PROGRAM MAIN
// =============================================================
// TEST RUCHU TRANSPORTEROW
// =============================================================
//
// Proba na maszynie: jedna paleta idzie trasa, w kazdym kroku
// pracuje PARA transporterow - ten, z ktorego paleta zjezdza,
// i ten, na ktory wjezdza.
//
// -------------------------------------------------------------
// CZUJNIKI
// -------------------------------------------------------------
// Podpiete czujniki koncza przejazd zamiast czasowki.
//
//   xUseSensors   = FALSE  wracamy na same czasowki, jak dotad
//   xStepWatchdog = FALSE  krok czeka na czujnik BEZ KONCA
//
// Na czas recznego wyzwalania czujnikow watchdog jest WYLACZONY:
// zaden krok nie przeskoczy sam, dopoki nie podasz sygnalu.
// Po podpieciu prawdziwych czujnikow warto go wlaczyc - wtedy
// martwy czujnik nie zatrzyma proby, tylko zglosi sie sam przez
// xStepTimeout i licznik nTimeouts.
//
// Kroki konczone czujnikiem:
//   st.2 -> st.3    IN2      st.7 -> st.8    IN7
//   st.3 -> st.4    IN3/IN4  st.8 -> st.11   IN8
//   st.6 -> st.7    IN5      st.12-> st.13   IN6
//   st.15-> st.16   IN10
//
// STACJA 1 nie ma czujnika w tej probie. Zamiast niego dziala
// bit xSt01_StackReady: TRUE = stoi tam stos i mozna nim jechac,
// zbocze 0 -> 1 = przyjechal nowy stos (licznik nStacksSeen).
//
// STACJA 4 bada JADACA palete - patrz ACT_MoveSt04.
//
// Wyjatkiem jest przejazd poprzeczny 8 -> 10: tam paleta lezy
// na lancuchu, rolki stacji 8 i 10 sa opuszczone i MUSZA stac.
// Jedzie sam falownik 7, przez tChainTime.
//
// -------------------------------------------------------------
// CO NIE JEST URUCHAMIANE
// -------------------------------------------------------------
// Falowniki 1, 2 i 3 sa ZABLOKOWANE w axDriveEnabled:
//   1  krzywka desztaplarki   - mechanika niegotowa
//   2  krzywka na stacji 8    - mechanika niegotowa
//   3  rolki dociskowe st. 4  - to nie jest transporter
//
// Blokada dziala niezaleznie od tabeli krokow: nawet gdyby
// krok zazadal takiego napedu, nie ruszy. Zeby go dopuscic,
// trzeba swiadomie ustawic bit w axDriveEnabled.
//
// -------------------------------------------------------------
// STEROWANIE
// -------------------------------------------------------------
//   START_TEST = TRUE   symulacja ruchu jedzie
//   START_TEST = FALSE  wszystkie napedy staja
//
//   xCmdResetDrives     kasuje bledy wszystkich falownikow,
//                       dziala na zbocze i sam sie zdejmuje
//
// Po wcisnieciu START maszyna sama sprawdza, czy ktorys naped
// nie stoi w bledzie, i probuje go skasowac - zanim cokolwiek
// ruszy. Jesli sie nie uda, zapala sie xResetFailed.
//
// Pelna aplikacja siedzi w PRG_Machine i na razie nie jest
// wywolywana.
VAR

	// =========================================================
	// STEROWANIE
	// =========================================================

	// GLOWNY BIT TESTU TRASY. TRUE = jedziemy, FALSE = stop.
	START_TEST			: BOOL;


	// =========================================================
	// PROBA CALOSCIOWA: DOWOZ -> DESZTAPLOWANIE -> STACJA 4
	// =========================================================
	//
	// Niezalezna od START_TEST. Wozi palety ze stacji 1 do
	// desztaplarki, potem kazda zwolniona palete przez stacje 4
	// z testem dociskow i ZATRZYMUJE ja na koncu stacji 4.
	// Palete zabiera sie stamtad recznie.

	// Potwierdzenie operatora: palety leza na stacji 1.
	// Kod sam go zdejmuje po przyjeciu - kolejny stos wymaga
	// podania go od nowa.
	xSt01_StackReady	: BOOL;

	// Start dowozu i obslugi transportu w tej probie
	START_FEED			: BOOL;

	// Ile palet przeszlo przez stacje 4
	nFeedPallets		: UDINT;

	// Podglad
	nFeedStep			: INT;
	sFeedPhase			: STRING(79);

	// Wewnetrzne sekwencji dowozu
	nFeedStepOld		: INT;
	xFeedNewStep		: BOOL;
	xFeedArmed			: BOOL;
	xFeedAdvance		: BOOL;
	tFeedStep			: TIME;
	tonFeedStep			: TON;
	rtrgFeedStart		: R_TRIG;

	// =========================================================
	// TOR WYJSCIOWY - DRUGA PALETA W MASZYNIE
	// =========================================================
	//
	// Transport jest rozbity na DWA niezalezne tory:
	//
	//   nFeedStep  tor A: stacja 1 -> 3 -> 4 -> cykl stacji 5
	//   nOutStep   tor B: stacja 5 -> 6 -> ... -> 16
	//
	// Dzieki temu paleta po rozrywaniu jedzie w strone stacji 16
	// SAMA, a desztaplarka moze w tym czasie wydac nastepna.
	// W maszynie sa wtedy dwie palety naraz.
	//
	// Zasob wspolny to transporter stacji 5 (naped 5) i blokada.
	// Dlatego tor A nie wjedzie na stacje 5, dopoki tor B z niej
	// nie zjedzie - patrz krok 75.
	//
	// nOutStep = 0 znaczy TOR B WOLNY.

	nOutStep			: INT;
	sOutPhase			: STRING(79);

	nOutStepOld			: INT;
	xOutNewStep			: BOOL;
	xOutArmed			: BOOL;
	xOutAdvance			: BOOL;
	tOutStep			: TIME;
	tonOutStep			: TON;

	// Stacja 5 skonczyla cykl i oddala palete torowi B.
	// Na tym sygnale desztaplarka wypuszcza nastepna palete.
	xSt05_Done			: BOOL;

	// Zadania startu torow. Tor URUCHAMIA SIE SAM, w swoim kroku 0.
	// Powod jest w komentarzu przy silniku krokow nizej - w skrocie:
	// krok wpisany z ZEWNATRZ wykonalby sie jeszcze w tym samym
	// cyklu, ze stara flaga xOutAdvance, i przeskoczylby natychmiast.
	// -----------------------------------------------------
	// STACJA 8 - POSADZENIE PALETY NOK NA LANCUCHU
	// -----------------------------------------------------
	//
	// Na stacji 8 nie ma blokady, a transporter chodzi tak
	// gladko, ze paleta zatrzymuje sie raz dalej, raz blizej.
	// Dlatego po tSt08_DropDelay od IN7 OPUSZCZAMY rolki: paleta
	// siada na lancuchu i to on ja wyhamowuje - zawsze tak samo.
	//
	// DOTYCZY WYLACZNIE PALET NOK, bo tylko one jada lancuchem.
	// Paleta OK jedzie dalej rolkami i zatrzymuje sie jak dotad -
	// dla niej nic sie nie zmienia.
	//
	// Dwie NIEZALEZNE czasowki od tego samego IN7:
	//   tFeedSt08Stop   zdjecie zadania z falownika (dobieg)
	//   tSt08_DropDelay opuszczenie rolek pod paleta
	tSt08_DropDelay		: TIME := T#830MS;
	tonSt08Drop			: TON;

	// Zatrzask: rolki stacji 8 maja zostac w dole, dopoki lancuch
	// nie zabierze palety. Bez niego kroki, ktore ich nie pisza,
	// podnosilyby je z powrotem.
	xSt08_RollDown		: BOOL;

	// Paleta jest na stacji 8 - od potwierdzenia IN7 do zabrania
	// jej przez lancuch. Na tej fladze chodzi tonSt08Drop, dzieki
	// czemu odliczanie NIE ZALEZY od tego, w ktorym kroku toru B2
	// paleta akurat stoi.
	xSt08_AtStation		: BOOL;

	// Czy TA paleta jedzie trasa odrzutu (lancuchem).
	// W tej probie wszystkie palety jada na stacje 16, wiec bit
	// jest TRUE. Gdy dojdzie klasyfikacja OK/NOK, ma go ustawiac
	// wynik badania, a nie operator.
	xSt08_PalletNOK		: BOOL := TRUE;

	xOutStart			: BOOL;
	xOut2Start			: BOOL;
	xOut3Start			: BOOL;

	// Droga ze stacji 5 wolna: tor B1 pusty i stacja 7 pusta
	xSt05_CanPass		: BOOL;

	// -----------------------------------------------------
	// BUFOROWANIE - TOR B ROZBITY NA TRZY ODCINKI
	// -----------------------------------------------------
	//
	// Odcinki wyznaczaja CZUJNIKI, bo tylko one wiedza, gdzie
	// naprawde stoi paleta:
	//
	//   nOutStep   B1  st.5 -> 6 -> 7    konczy sie na IN5
	//   nOut2Step  B2  st.7 -> 8         konczy sie na IN7
	//   nOut3Step  B3  st.8 -> ... -> 16 konczy sie na IN10
	//
	// Kazdy odcinek zwalnia sie DOPIERO wtedy, gdy nastepny
	// przejmie palete. Dzieki temu w obiegu moga byc naraz:
	// paleta na stacji 5, paleta na 7, paleta na 8 i paleta
	// w drodze na 16 - zamiast jednej na cala maszyne.
	//
	// Transporter stacji 7 (naped 11) obsluguje B1 i B2, a rolki
	// stacji 8 (naped 12) B2. Dlatego paleta czeka w krokach
	// 205 i 218 z ZATRZYMANYMI napedami, zamiast dojezdzac
	// wprost na zajety odcinek.

	nOut2Step			: INT;
	sOut2Phase			: STRING(79);
	nOut2StepOld		: INT;
	xOut2NewStep		: BOOL;
	xOut2Armed			: BOOL;
	xOut2Advance		: BOOL;
	tOut2Step			: TIME;
	tonOut2Step			: TON;

	nOut3Step			: INT;
	sOut3Phase			: STRING(79);
	nOut3StepOld		: INT;
	xOut3NewStep		: BOOL;
	xOut3Armed			: BOOL;
	xOut3Advance		: BOOL;
	tOut3Step			: TIME;
	tonOut3Step			: TON;

	// -----------------------------------------------------
	// STACJA 5 - CZAS PCHANIA PALETY DO BLOKADY
	// -----------------------------------------------------
	//
	// Paleta opiera sie o blokade duzo wczesniej, niz konczy sie
	// krok 80. Kazda sekunda ponad to jest transporterem
	// mielacym pod stojaca paleta - tak przeciazamy naped 5.
	// Po tym czasie napedy 4 i 5 STAJA, a krok trwa dalej.
	//
	// DOMYSLNIE ROWNE tFeedToSt05 - czyli tak, jak bylo przed
	// wprowadzeniem tej nastawy. Moje 4 s bylo za krotkie
	// i paleta nie dojezdzala do blokady.
	//
	// Skracaj DOPIERO po obejrzeniu, gdzie paleta sie zatrzymuje:
	// ma byc na tyle dlugie, zeby doszla do blokady, i na tyle
	// krotkie, zeby transporter nie mielil pod nia bez potrzeby.
	tSt05_Push			: TIME := T#9S;
	tonSt05Push			: TON;

	// -----------------------------------------------------
	// STACJA 4 - ROLKI DOCISKOWE (NAPED 3)
	// -----------------------------------------------------
	//
	// Kreca sie razem z transporterem stacji 4 (naped 4).
	// Bit ponizej wybiera kierunek obrotu - do ustawienia
	// online, bez pobierania projektu.
	xSt04_RollRev		: BOOL := TRUE;

	// Stan dociskow stacji 4 w tej probie - przepisywany co cykl
	xFeedPressOn		: BOOL;
	xFeedPressLoOn		: BOOL;

	// Czas przejazdu st.4 -> st.5. Stacja 5 nie ma czujnika,
	// wiec dojazd konczy sie czasowka. Dobrane na maszynie.
	tFeedToSt05			: TIME := T#9S;

	// DOBIEG NA STACJI 3. Czujnik IN2 widzi krawedz natarcia
	// stosu, a szczeki maja trafic pod DRUGA palete od dolu -
	// stos musi wiec dojechac jeszcze kawalek po wykryciu.
	//
	// ZERO = stop natychmiast po czujniku, czyli tak, jak bylo.
	// Odpowiednik tSt04_StopDelay dla stacji 4.
	tFeedSt03Stop		: TIME := T#0S;

	// Odstep od zatrzymania palety na stacji 5 do ruszenia
	// mechaniki. Stacja 5 nie ma czujnika, wiec nie wiemy, kiedy
	// paleta oprze sie o blokade - dajemy jej na to czas.
	tSt05_Settle		: TIME := T#8S;

	// Stan mechaniki stacji 5 w tej probie - kazdy krok podaje
	// swoj pelny stan, cewki przepisujemy co cykl.
	xFeed05_Block		: BOOL;		// blokada wysunieta
	xFeed05_Lift		: BOOL;		// szczeki podniesione
	xFeed05_Jaws		: BOOL;		// szczeki zamkniete
	xFeed05_Pull		: BOOL;		// silowniki rozrywajace w gorze

	// Diagnostyka napedow zadanych przez biezacy krok
	nFeedBadDrv			: INT;
	sFeedDrvWhy			: STRING(31);
	tonFeedDrv			: TON;

	// -----------------------------------------------------
	// CZASOWKI PRZEJAZDOW BEZ CZUJNIKA
	// -----------------------------------------------------
	//
	// Odcinki, na ktorych nie ma czym potwierdzic dojazdu.
	// Tam, gdzie czujnik jest, czasowka nie jest uzywana wcale.

	tFeed5to6			: TIME := T#12S;		// st.5 -> st.6
	tFeed9Chain			: TIME := T#19S;		// lancuch st.8 -> st.10
	tFeed10to14			: TIME := T#8S;		// st.10 -> st.14
	tFeed14to15			: TIME := T#8S;		// st.14 -> st.15

	// Paleta zniknela z czujnika stacji 16. Po tym czasie
	// uznajemy stacje za pusta - odbiera ja operator.
	tSt16_Clear			: TIME := T#4S;

	// -----------------------------------------------------
	// DOBIEGI PO CZUJNIKACH
	// -----------------------------------------------------
	//
	// Czujnik widzi krawedz natarcia palety, a ona ma stanac
	// na srodku stacji. ZERO = stop natychmiast po czujniku.
	// Odpowiedniki tFeedSt03Stop i tSt04_StopDelay.

	tFeedSt08Stop		: TIME := T#740MS;		// IN7  stacja 8
	tFeedSt16Stop		: TIME := T#0S;		// IN10 stacja 16

	// Rolki podnoszone stacji 8 i 10. TRUE = w gorze, czyli
	// transport wzdluz. Na czas przejazdu lancuchem OBIE musza
	// zejsc, inaczej szarpalyby palete z dwoch stron.
	xFeedRoll08Up		: BOOL := TRUE;
	xFeedRoll10Up		: BOOL := TRUE;

	// Zezwolenie z lancucha bezpieczenstwa
	xSafetyOK			: BOOL := TRUE;

	// KASOWANIE BLEDOW WSZYSTKICH FALOWNIKOW - dziala na zbocze.
	// Bit sam sie zdejmuje po wystawieniu impulsu.
	xCmdResetDrives		: BOOL;

	// Automatyczne kasowanie bledow po wcisnieciu START.
	// FALSE = start nie probuje niczego kasowac.
	xAutoResetOnStart	: BOOL := TRUE;

	// Odstep miedzy kolejnymi probami kasowania
	tResetGap			: TIME := T#1S;

	// Czestotliwosc BAZOWA transporterow [Hz]. Uzywana wszedzie,
	// gdzie alrDriveFreq nie ma wpisanej wlasnej wartosci.
	lrTestFreq			: LREAL := 20.0;

	// =========================================================
	// CZESTOTLIWOSC OSOBNO DLA KAZDEGO NAPEDU [Hz]
	// =========================================================
	//
	// Zero znaczy "uzyj lrTestFreq". Wpisanie liczby dotyczy
	// tylko tego jednego falownika.
	//
	// Przydzial stacja -> falownik:
	//   st.1  -> 8     st.5  -> 5     st.9  -> 7      st.13 -> 15
	//   st.2  -> 9     st.6  -> 6     st.10 -> 16     st.14 -> 17
	//   st.3  -> 10    st.7  -> 11    st.11 -> 13     st.15 -> 18
	//   st.4  -> 4     st.8  -> 12    st.12 -> 14     st.16 -> 19
	//
	// Krzywki 1 i 2 maja wlasna lrCamFreq i ta tablica ich nie
	// dotyczy.
	//
	// UWAGA: naped czyta czestotliwosc przy STARCIE (M_Start jest
	// wolane na zboczu). Zmiana w trakcie jazdy zadziala dopiero
	// przy nastepnym ruszeniu.

	alrDriveFreq		: ARRAY[1..20] OF LREAL;

	// Czas jednego kroku - przejazd palety miedzy stacjami
	tStepTime			: TIME := T#5S;

	// Przejazd poprzeczny transporterem lancuchowym jest dluzszy
	tChainTime			: TIME := T#6S;

	// Czas jednego ruchu silownika. Czujnikow polozenia jeszcze
	// nie ma, wiec po tym czasie uznajemy ruch za wykonany.
	tCylTime			: TIME := T#2S;

	// Stacja 4 - dociski gorne i dolne maja isc praktycznie razem.
	// Gorne schodza pierwsze, dolne po tym krotkim odstepie,
	// zeby dolne nie uniosly palety. Cofanie jest jednoczesne.
	tSt04_UpToLo		: TIME := T#2200MS;

	// FALSE = same transportery, silowniki stoja
	xCylEnable			: BOOL := TRUE;


	// =========================================================
	// CZUJNIKI
	// =========================================================
	//
	// FALSE = jedziemy na samych czasowkach, tak jak dotad.
	// TRUE  = kroki wypisane w ACT_Move koncza sie czujnikiem,
	//         a czasowka pracuje juz tylko jako watchdog.

	xUseSensors			: BOOL := TRUE;

	// STACJA 1 - czujnika IN1 NIE uzywamy. Zastepuje go bit
	// xSt01_StackReady zadeklarowany na gorze.
	nStacksSeen			: UDINT;

	// Obraz czujnikow sprowadzony do JEDNEGO znaczenia:
	// TRUE = PALETA JEST. Polaryzacje ustawia ACT_Inputs i tylko on.
	xPal_St03			: BOOL;		// IN2   stacja 3
	xPal_St04In			: BOOL;		// IN3   wjazd na stacje 4
	xPal_St04End		: BOOL;		// IN4   koniec testu desek
	xPal_St07			: BOOL;		// IN5   stacja 7
	xPal_St13			: BOOL;		// IN6   koniec stacji 13
	xPal_St08			: BOOL;		// IN7   stacja 8
	xPal_St11			: BOOL;		// IN8   stacja 11
	xPal_St16			: BOOL;		// IN10  stacja 16

	// Surowe wejscia - do podgladu bez otwierania GVL
	axInRaw				: ARRAY[1..10] OF BOOL;

	// -----------------------------------------------------
	// POLARYZACJA CZUJNIKOW - JEDYNE MIEJSCE
	// -----------------------------------------------------
	//
	// TRUE  = czujnik ROZWIERA przy palecie (0 = paleta)
	// FALSE = czujnik ZWIERA przy palecie   (1 = paleta)
	//
	// Wartosci ponizej sa wg opisu z maszyny. Jesli ktorys
	// czujnik zachowa sie odwrotnie, przestawia sie JEDEN bit
	// online - bez zmiany kodu i bez pobierania projektu.
	//
	//   1  st.1              nieuzywany
	//   2  st.3              ROZWIERA - stwierdzone na maszynie,
	//                        wbrew pierwotnemu opisu
	//   3  wjazd st.4        rozwiera
	//   4  koniec testu st.4 rozwiera
	//   5  st.7              zwiera
	//   6  koniec st.13      rozwiera
	//   7  st.8              zwiera
	//   8  st.11             zwiera
	//   9  niepodlaczony
	//  10  st.16             zwiera

	axInInverted		: ARRAY[1..10] OF BOOL :=
	                      [FALSE, TRUE, TRUE, TRUE, FALSE,
	                       TRUE, FALSE, FALSE, FALSE, FALSE];

	// WATCHDOG KROKU CZUJNIKOWEGO.
	//
	// FALSE = krok czeka na czujnik BEZ KONCA. Tak jedziemy przy
	//         recznym wyzwalaniu czujnikow - nic nie przeskoczy
	//         kroku, dopoki sam nie podasz sygnalu.
	// TRUE  = po tMoveTimeout krok konczy sie mimo wszystko,
	//         zapala sie xStepTimeout i rosnie nTimeouts.
	xStepWatchdog		: BOOL := FALSE;

	tMoveTimeout		: TIME := T#20S;
	xStepTimeout		: BOOL;
	nTimeouts			: UDINT;


	// =========================================================
	// STACJA 4 - TEST NA JADACEJ PALECIE
	// =========================================================
	//
	// Paleta nie zatrzymuje sie pod rolkami. Czujnik wjazdu (IN3)
	// odlicza tSt04_EntryToPress i wtedy rolki schodza na deski.
	// Czujnik konca testu (IN4) NATYCHMIAST je cofa, a transporter
	// stoi tSt04_StopDelay pozniej - paleta dojezdza do konca stacji.

	tSt04_EntryToPress	: TIME := T#2600MS;
	tSt04_StopDelay		: TIME := T#300MS;


	// =========================================================
	// SZTAPLARKA I DESZTAPLARKA
	// =========================================================
	//
	// Dwa NIEZALEZNE cykle, kazdy z wlasnym bitem startu. Nie
	// maja nic wspolnego z START_TEST.
	//
	// Poziom TRUE = cykl pracuje.
	// Poziom FALSE = natychmiastowy stop, hamulec zaklada sie
	//                tCamBrakeHold pozniej.
	//
	// REGULA NADRZEDNA obu maszyn: nic w szczekach = szczeki
	// OTWARTE i jazda na pozycje DOLNA, niezaleznie od tego,
	// gdzie wozek stoi. Cykl zaczyna sie i konczy na dole
	// z otwartymi szczekami.

	START_DESTACK		: BOOL;		// desztaplarka, stacja 3
	START_STACK			: BOOL;		// sztaplarka, stacja 11

	// -----------------------------------------------------
	// JAZDA RECZNA KRZYWKA
	// -----------------------------------------------------
	//
	// Trzymasz bit - wozek jedzie. Puszczasz - staje, hamulec
	// zaklada sie tCamBrakeHold pozniej, tak samo jak w cyklu.
	//
	// Dziala TYLKO przy zdjetym starcie danej maszyny, zeby
	// nigdy nie walczyc z sekwencja. Sluzy do sprawdzenia,
	// czy enkoder liczy i w ktora strone.

	JOG_DESTACK_FWD		: BOOL;
	JOG_DESTACK_REV		: BOOL;
	JOG_STACK_FWD		: BOOL;
	JOG_STACK_REV		: BOOL;

	xDeJog				: BOOL;
	xStJog				: BOOL;

	// -----------------------------------------------------
	// UCZENIE POZYCJI
	// -----------------------------------------------------
	//
	// Dojedz jogiem tam, gdzie wozek ma stawac, i podaj bit.
	// Zbocze 0 -> 1 przepisuje BIEZACA pozycje enkodera do
	// odpowiedniej nastawy. Koniec z wpisywaniem liczb z palca.
	//
	// UWAGA: nastawy siedza na razie w MAIN, wiec pobranie
	// projektu je kasuje. Po ustaleniu przenosimy do GVL_PERSIST.

	TEACH_DE_BOTTOM		: BOOL;
	TEACH_DE_MIDDLE		: BOOL;
	TEACH_DE_TOP		: BOOL;
	TEACH_ST_BOTTOM		: BOOL;
	TEACH_ST_MIDDLE		: BOOL;
	TEACH_ST_TOP		: BOOL;

	rtrgTeach			: ARRAY[1..6] OF R_TRIG;

	// Ostatnio nauczona pozycja - potwierdzenie na podgladzie
	sTeachLast			: STRING(79);

	// Czestotliwosc krzywek. Osobno od transporterow.
	// Nizej niz transportery - wolniej znaczy krotszy dojazd
	// po zdjeciu zadania, a wiec mniejszy blad pozycji.
	lrCamFreq			: LREAL := 15.0;

	// Ruch szczek - czujnikow polozenia nie ma
	tJawTime			: TIME := T#2S;


	// Odstep od ZALOZENIA hamulca do chwytu szczekami.
	// Wozek musi sie uspokoic, zanim szczeki wejda pod palete.
	tDeGripDelay		: TIME := T#1S;

	// -----------------------------------------------------
	// POZYCJE I LICZNIKI SIEDZA W GVL_PERSIST
	// -----------------------------------------------------
	//
	// Nastawy:  GVL_PERSIST.St03.Cfg.diPosBottom / Middle / Top
	//           GVL_PERSIST.St11.Cfg.diPosBottom / Middle / Top
	//           GVL_PERSIST.St03.Cfg.nStackSize
	// Liczniki: GVL_PERSIST.St03.Mem.nRemaining / nHeld
	//           GVL_PERSIST.St11.Mem.nHeld
	//
	// Sa NIEULOTNE, wiec przezywaja zanik zasilania, aktywacje
	// konfiguracji i reset cold. Uczenie pozycji zapisuje wprost
	// tam - nie ma drugiej kopii, ktora moglaby sie rozjechac.



	// Wyprzedzenie hamowania - zadanie znika tyle przed celem.
	// Zaczynamy od zera i ustawiamy z odczytu diCoast.
	diCamStopLead		: DINT := 0;

	// Okno "jestem na miejscu" przy bazowaniu. Bez niego wozek
	// stojacy tuz przy dolnej pozycji robilby caly obrot, zeby
	// do niej "dojechac".
	diCamTol			: DINT := 300;

	// Ile impulsow za celem uznajemy jeszcze za "jestem".
	// Musi byc WIEKSZE niz dojazd po zdjeciu zadania, inaczej
	// wozek stojacy tuz ZA punktem objechalby caly obrot,
	// zeby do niego wrocic.
	diCamOvershoot		: DINT := 5000;

	// -----------------------------------------------------
	// DOKAD JEDZIE BIEZACY KROK
	// -----------------------------------------------------
	//
	// Krok podaje WARTOSC ENKODERA, do ktorej ma dojechac,
	// a droge liczymy raz, przy wejsciu w krok, z zywej
	// pozycji. Nigdzie nie zakladamy, ile impulsow ma cykl
	// maszyny - to bylo zrodlo kumulujacego sie bledu.

	diDeGoToEnc			: DINT;
	diStGoToEnc			: DINT;

	// -----------------------------------------------------
	// POMIAR - ILE IMPULSOW MA NAPRAWDE CYKL MASZYNY
	// -----------------------------------------------------
	//
	// diDeCycleCounts   droga przejechana miedzy kolejnymi
	//                   dolnymi pozycjami. Jesli enkoder jest
	//                   1:1 z korba, ma byc okolo 65536.
	//                   Kazda inna liczba znaczy, ze cykl
	//                   maszyny to nie jest jeden obrot enkodera.
	// diDeBottomErr     o ile minelismy nauczony dol, ze znakiem
	// diDeCoastMax      najwiekszy zaobserwowany dojazd. Musi
	//                   byc MNIEJSZY niz diCamOvershoot, inaczej
	//                   ruch do punktu tuz za nami pojedzie
	//                   dookola.

	diDeCycleCounts		: DINT;
	diDeBottomErr		: DINT;
	diDeCoastMax		: DINT;

	diStCycleCounts		: DINT;
	diStBottomErr		: DINT;
	diStCoastMax		: DINT;

	// Ustawienie punktu odniesienia osi, impuls jednocyklowy
	xDeSetAccum			: BOOL;
	xStSetAccum			: BOOL;
	diDeAccumSet		: DINT;
	diStAccumSet		: DINT;

	// Roboczy
	diTmp				: DINT;

	// -----------------------------------------------------
	// KONTROLA POPRAWNOSCI NASTAW POZYCJI
	// -----------------------------------------------------
	//
	// Trzy pozycje musza byc od siebie ODDALONE. Zerowe albo
	// pomylone nastawy oznaczaja, ze wozek "juz jest na miejscu"
	// w kazdym kroku - a wtedy szczeki zamykaja sie na dole,
	// na stosie. Cykl nie ma prawa ruszyc na takich nastawach.

	xDeCfgOK			: BOOL;
	xStCfgOK			: BOOL;
	diCamMinSpan		: DINT := 1000;

	// -----------------------------------------------------
	// KONTROLA ENKODERA PO STARCIE
	// -----------------------------------------------------
	//
	// Enkoder absolutny powinien utrzymac wartosc przez zanik
	// zasilania. Zapamietujemy ja na biezaco w GVL_PERSIST
	// i po starcie porownujemy z odczytem. Zgadza sie -
	// bazowanie jest zbedne. Nie zgadza sie - kod to zglasza,
	// zamiast po cichu jechac wedlug zlych pozycji.

	xEncCheckDone		: BOOL;
	diDeEncJump			: DINT;
	diStEncJump			: DINT;
	sEncCheck			: STRING(79);

	// Ile impulsow roznicy jeszcze wybaczamy po starcie
	diEncCheckTol		: DINT := 500;

	// START: wyprzedzenie zdjecia hamulca przed komenda dla
	// falownika. ZERO = jednoczesnie, i tak ma byc.
	tCamBrakeRelease	: TIME := T#0S;

	// STOP: ile hamulec czeka po zdjeciu komendy z falownika.
	// Rampa hamowania falownika to 1 s, wiec hamulec zaciska sie
	// na wolno obracajacym sie jeszcze wale - SWIADOMIE, zeby
	// nie puszczac wozka wolno.
	tCamBrakeHold		: TIME := T#700MS;

	// Kasowanie czuwaka obu osi, dziala na zbocze
	RESET_CAM			: BOOL;

	// =========================================================
	// RESET CYKLU DO ZERA
	// =========================================================
	//
	// Po recznym oproznieniu maszyny z palet. Sprowadza obie
	// maszyny i transport do kroku 0, zeruje liczniki palet
	// i uzgodnienia, kasuje czuwaki osi.
	//
	// NICZYM NIE RUSZA. Wozki wroca na dol dopiero przy starcie,
	// bo krok 0 obu maszyn to "szczeki otwarte, jazda na dol".
	//
	// Bit sam sie zdejmuje.

	RESET_CYCLE			: BOOL;
	rtrgResetCycle		: R_TRIG;

	// -----------------------------------------------------
	// PODGLAD OSI
	// -----------------------------------------------------

	fbCamDestack		: FB_CamAxis;
	fbCamStack			: FB_CamAxis;

	nDeStep				: INT;
	nStStep				: INT;
	sDePhase			: STRING(79);
	sStPhase			: STRING(79);
	nDeCycles			: UDINT;
	nStCycles			: UDINT;

	// -----------------------------------------------------
	// LICZNIKI PALET
	// -----------------------------------------------------
	//
	// GVL_PERSIST.St03.Mem.nRemaining  ile palet zostalo w desztaplarce razem:
	//               na transporterze plus wiszace na szczekach
	// GVL_PERSIST.St03.Mem.nHeld       ile wisi na szczekach desztaplarki
	// GVL_PERSIST.St11.Mem.nHeld       ile palet liczy stos w sztaplarce


	// -----------------------------------------------------
	// UZGODNIENIA Z TRANSPORTEM
	// -----------------------------------------------------

	// Desztaplarka zwolnila palete - transport moze ja zabrac
	xDe_PalletReleased	: BOOL;

	// Desztaplarka pusta, cykl zamkniety na pozycji dolnej
	xDe_Empty			: BOOL;

	// Sztaplarka ma pelny stos na transporterze
	xSt_StackReady		: BOOL;

	// -----------------------------------------------------
	// CZASOWKI OD ZALOZENIA HAMULCA
	// -----------------------------------------------------
	//
	// Licza dopiero od chwili, w ktorej hamulec sie ZACISNIE -
	// nie od wejscia w krok.

	tonDeBrake			: TON;
	tonStBrake			: TON;
	tDeBrakeWait		: TIME;
	tStBrakeWait		: TIME;

	// Czujnik musi byc najpierw WOLNY, zeby sie zaliczyl
	xDeArmed			: BOOL;
	xStArmed			: BOOL;

	// Stan szczek deklarowany przez KAZDY krok i przepisywany
	// na cewki co cykl. Poleganie na tym, ze cewka zachowa
	// wartosc miedzy krokami, juz raz nas kosztowalo prawdziwy
	// blad - ACT_ClearCoils zeruje je w kazdym cyklu.
	xDeJawsClosed		: BOOL;
	xStJawsClosed		: BOOL;

	// -----------------------------------------------------
	// ZYCIE ENKODEROW
	// -----------------------------------------------------
	//
	// Rosna przy KAZDEJ zmianie pozycji. Jesli silnik chodzi,
	// a licznik stoi - enkoder nie jest podlinkowany albo nie
	// liczy. To rozstrzyga sprawe w jednej liczbie.

	nDeEncMoves			: UDINT;
	nStEncMoves			: UDINT;
	diDePosOld			: DINT;
	diStPosOld			: DINT;

	tonDeStep			: TON;
	tonStStep			: TON;
	xDeAdvance			: BOOL;
	xStAdvance			: BOOL;
	tDeStep				: TIME;
	tStStep				: TIME;

	// Zadanie dla osi - liczone przez maszyne stanow,
	// podawane do bloku JEDNYM wywolaniem na cykl
	xDeGo				: BOOL;
	xStGo				: BOOL;
	diDeTarget			: DINT;
	diStTarget			: DINT;

	// Wykrycie zmiany kroku. Bez tego krok zaliczylby xInPos
	// z POPRZEDNIEJ pozycji i przeskoczyl dwa kroki naraz.
	nDeStepOld			: INT;
	nStStepOld			: INT;
	xDeNewStep			: BOOL;
	xStNewStep			: BOOL;
	xDeAtPos			: BOOL;
	xStAtPos			: BOOL;

	rtrgDeStart			: R_TRIG;
	rtrgStStart			: R_TRIG;

	// Cewki hamulcow. TRUE = hamulec ROZLACZONY.
	xBrakeDestack		: BOOL;
	xBrakeStack			: BOOL;


	// =========================================================
	// RECZNE STEROWANIE POJEDYNCZYM SILOWNIKIEM
	// =========================================================
	//
	// Do sprawdzenia okablowania bez sekwencji. Gdy nManCyl <> 0,
	// sekwencja stoi, transportery stoja, a wybrany silownik
	// slucha bitow ponizej.
	//
	//    1  st.3  szczeki desztaplarki
	//    2  st.4  dociski gorne
	//    3  st.4  dociski dolne
	//    4  st.5  blokada
	//    5  st.5  podnoszenie szczek
	//    6  st.5  szczeki (zamkniecie / otwarcie)
	//    7..12 st.5 silowniki rozrywajace 1..6
	//   13  st.8  rolki podnoszone
	//   14  st.10 rolki podnoszone
	//   15  st.11 szczeki sztaplarki

	nManCyl				: INT;
	xManExtend			: BOOL;
	xManRetract			: BOOL;


	// =========================================================
	// DOPUSZCZENIE NAPEDOW
	// =========================================================
	//
	// FALSE = naped nie ruszy, chocby krok tego zadal.
	// Ustawiane w ACT_Config, mozna zmieniac online.

	axDriveEnabled		: ARRAY[1..20] OF BOOL;


	// =========================================================
	// KIERUNEK OBROTOW
	// =========================================================
	//
	// TRUE = jazda w druga strone. Silniki stacji 1, 5, 6, 7,
	// 8, 9, 14, 15, 16 sa podlaczone odwrotnie - do poprawy
	// w szafie, na razie odwracamy bit.

	axReverse			: ARRAY[1..20] OF BOOL;


	// =========================================================
	// PODGLAD
	// =========================================================

	// Gdzie jest wirtualna paleta i co sie z nia dzieje
	nIdx				: INT;		// pozycja na trasie
	nSub				: INT;		// krok sekwencji stacji
	xMoving				: BOOL;		// TRUE = przejazd, FALSE = praca stacji
	sPhase				: STRING(79);

	// Ktore napedy maja teraz pracowac
	axRunReq			: ARRAY[1..20] OF BOOL;

	// Stan napedow
	aeDrvState			: ARRAY[1..20] OF E_NordSK550P_State;
	axDrvRunning		: ARRAY[1..20] OF BOOL;
	alrDrvFreqAct		: ARRAY[1..20] OF LREAL;

	// UWAGA - to sa DWIE ROZNE rzeczy:
	//   axDrvFault  blad zglaszany przez falownik (bit 3 StatusWord)
	//   axDrvError  jakakolwiek blokada: blad, brak zezwolenia
	//               albo zerwana komunikacja
	axDrvFault			: ARRAY[1..20] OF BOOL;
	axDrvError			: ARRAY[1..20] OF BOOL;

	// Slowa sterujace i statusowe - do czytania, co naped
	// naprawde zglasza
	awDrvStatus			: ARRAY[1..20] OF UINT;
	awDrvControl		: ARRAY[1..20] OF UINT;

	// Ktorykolwiek naped zglasza blad
	xAnyDriveError		: BOOL;
	xAnyDriveFault		: BOOL;

	// Kasowanie nie poskutkowalo - blad wraca albo trzyma
	xResetFailed		: BOOL;

	// Trwa kasowanie bledow przed startem
	xResetInProgress	: BOOL;
	nResetTries			: INT;

	// Blokada zadzialala - lancuch wymusil postoj rolek 8 i 10
	xChainInterlock		: BOOL;

	// Blokada stacji 5 kontra transporter - patrz ACT_ApplyDrives
	xSt05_BlockLock		: BOOL;
	tonSt05BlockDown	: TON;

	// Czas biezacego kroku
	tThisStep			: TIME;

	// Licznik pelnych przebiegow trasy
	nLoops				: UDINT;

	// =========================================================
	// LICZNIKI ZYCIA - do sprawdzenia, co sie naprawde wykonuje
	// =========================================================
	//
	// nCycles     rosnie w kazdym cyklu zadania. Jesli stoi,
	//             MAIN sie nie wykonuje albo wysypal sie wczesniej.
	// nOutWrites  rosnie za kazdym przepisaniem cewek na wyjscia.
	//             Jesli nCycles rosnie, a nOutWrites stoi -
	//             program nie dochodzi do ACT_Outputs.
	// nCoilsOn    ile cewek jest w tej chwili podanych. Jesli
	//             rosnie i spada, a nic sie nie rusza - sygnal
	//             nie dochodzi do zaworu.

	nCycles				: UDINT;
	nOutWrites			: UDINT;
	nCoilsOn			: INT;


	// =========================================================
	// CEWKI ZAWOROW
	// =========================================================
	//
	// Stan trzymany miedzy cyklami. ACT_Outputs przepisuje go
	// na wyjscia - mapowanie jest TAM i tylko tam.

	// Stacja 3 - szczeki desztaplarki
	xSt03_JawClose		: BOOL;
	xSt03_JawOpen		: BOOL;

	// Stacja 4 - dociski. Obie grupy gornych chodza razem.
	xSt04_UpExt			: BOOL;
	xSt04_UpRet			: BOOL;
	xSt04_LoExt			: BOOL;
	xSt04_LoRet			: BOOL;

	// Stacja 5
	xSt05_BlockExt		: BOOL;		// blokada wysuw
	xSt05_BlockRet		: BOOL;		// blokada opuszczenie
	xSt05_LiftUp		: BOOL;		// szczeki w gore
	xSt05_LiftDown		: BOOL;		// szczeki w dol
	xSt05_JawClose		: BOOL;		// trzy pary szczek razem
	axSt05_PullUp		: ARRAY[1..6] OF BOOL;
	axSt05_PullDown		: ARRAY[1..6] OF BOOL;

	// Rolki podnoszone
	xSt08_Up			: BOOL;
	xSt08_Down			: BOOL;
	xSt10_Up			: BOOL;
	xSt10_Down			: BOOL;

	// Stacja 11 - szczeki sztaplarki
	xSt11_JawClose		: BOOL;
	xSt11_JawOpen		: BOOL;


	// =========================================================
	// NAPEDY
	// =========================================================

	fbNord				: ARRAY[1..20] OF FB_NordSK550PP;


	// =========================================================
	// OBSERWATOR STANU - LOG CSV NA DYSKU STEROWNIKA
	// =========================================================
	//
	// Co tLogPeriod jeden wiersz z kluczowymi zmiennymi, a do
	// tego wiersz na kazde ZDARZENIE: zmiana numeru kroku,
	// czujnika, zadania napedu, bledu falownika, bitu operatora,
	// szczek, skok enkodera. Najwyzej jeden wiersz na cykl.
	//
	// Nowy plik: start PLC, RESET_CYCLE, zbocze xLogNewFile.
	// Katalog MUSI istniec na sterowniku: fbLog.sDir
	// (domyslnie C:\TesterPalet\log\). Nazwa pliku w fbLog.sFileName.
	//
	// Logger tylko CZYTA zmienne procesu - ACT_Logger idzie jako
	// ostatnia akcja cyklu, po ACT_Outputs, zeby w pliku bylo to,
	// co naprawde poszlo na wyjscia.

	fbLog				: FB_CsvLogger;

	// FALSE = nie zbieramy wierszy (plik zostaje, nic sie nie psuje)
	xLogEnable			: BOOL := TRUE;

	// Zbocze = nowy plik bez resetu cyklu. Sam sie zdejmuje.
	xLogNewFile			: BOOL;

	// Takt wiersza okresowego
	tLogPeriod			: TIME := T#1S;
	tonLog				: TON;

	// Skok enkodera w jednym cyklu, od ktorego piszemy zdarzenie
	diLogEncJump		: DINT := 2000;

	// Powod biezacego wiersza - do kolumny "why"
	sLogWhy				: STRING(79);
	xLogEvent			: BOOL;
	nLogRows			: UDINT;

	// Pamiec do wykrywania zdarzen
	xLogInit			: BOOL;
	anLogStepOld		: ARRAY[1..6] OF INT;
	axLogInOld			: ARRAY[1..10] OF BOOL;
	axLogReqOld			: ARRAY[1..20] OF BOOL;
	axLogFaultOld		: ARRAY[1..20] OF BOOL;
	axLogBitOld			: ARRAY[1..24] OF BOOL;
	axLogBit			: ARRAY[1..24] OF BOOL;

	// Robocze do skladania nazw kolumn napedow
	sLogPfx				: STRING(15);
	wLogFesto1			: WORD;
	wLogFesto2			: WORD;
	nLogI				: INT;
	nLogJ				: INT;


	// =========================================================
	// WEWNETRZNE
	// =========================================================

	xInit				: BOOL;
	i					: INT;
	lrThisFreq			: LREAL;
	tonStep				: TON;
	tonResetGap			: TON;
	xAdvance			: BOOL;
	rtrgStart			: R_TRIG;
	rtrgResetDrv		: R_TRIG;
	rtrgStack			: R_TRIG;
	xDoResetPulse		: BOOL;
	axRunOld			: ARRAY[1..20] OF BOOL;

	// Krok zglasza tu, ze czeka na czujnik i ktory to czujnik.
	// Kasowane co cykl, ustawiane przez sam krok.
	xWaitSensor			: BOOL;
	xSensorOK			: BOOL;

	// Czujnik musi najpierw byc WOLNY. Bez tego zaliczylby sie
	// stan sprzed kroku albo czujnik zawieszony na stale.
	xStepArmed			: BOOL;

	// Wykrycie zmiany kroku - czasowka i uzbrojenie od zera
	xNewStep			: BOOL;
	nIdxOld				: INT;
	nSubOld				: INT;
	xMovingOld			: BOOL;

	// TRUE = przejazd ma jeszcze kroki wewnetrzne, nIdx zostaje
	xHoldIdx			: BOOL;

END_VAR
VAR CONSTANT

	// P105 falownikow
	cFmax				: LREAL := 50.0;

	// Liczba falownikow zmapowanych w .tsproj
	cNumDrives			: INT := 19;

	// Liczba pozycji na trasie
	cLastIdx			: INT := 16;

	// Ile razy probujemy skasowac blad przed startem
	cResetTries			: INT := 3;

END_VAR

// =============================================================
// MAIN - TEST RUCHU TRANSPORTEROW
// =============================================================

// Puls zycia - jesli ten licznik stoi, MAIN sie nie wykonuje
nCycles := nCycles + 1;

ACT_Config();

ACT_Inputs();

ACT_Sequence();

// Krzywki chodza NIEZALEZNIE od START_TEST i po ACT_Sequence,
// zeby ich szczeki mialy pierwszenstwo przed sekwencja linii.
ACT_CamCycles();

// Transport proby calosciowej - po krzywkach, zeby jego
// cewki i zadania napedow mialy pierwszenstwo.
ACT_TestFeed();

ACT_ResetDrives();

ACT_ApplyDrives();

ACT_Drives();

ACT_Outputs();

// Obserwator stanu - OSTATNI, zeby logowal to, co poszlo na wyjscia
ACT_Logger();

ACTION ACT_ApplyDrives:
// =============================================================
// ACT_ApplyDrives
// Zadanie ruchu -> metody falownikow
// =============================================================
//
// Metody wolamy NA ZBOCZU. Blok napedu przy blokadzie sam kasuje
// zadanie ruchu i naped nie moze ruszyc sam po ustapieniu
// przyczyny - wolanie M_Start co cykl zepsuloby to zabezpieczenie.

xAnyDriveError := FALSE;


// -------------------------------------------------------------
// BLOKADA: LANCUCH KONTRA ROLKI STACJI 8 I 10
// -------------------------------------------------------------
//
// Gdy jedzie transporter lancuchowy, rolki stacji 8 i 10 sa
// opuszczone i paleta lezy na lancuchu. Krecenie nimi w tym
// czasie szarpaloby palete z dwoch stron naraz.
//
// To nie jest poprawka tabeli krokow, tylko warunek nadrzedny -
// zadziala takze wtedy, gdy ktos pozniej zmieni tabele.

xChainInterlock := FALSE;

IF axRunReq[7] THEN

	IF axRunReq[12] OR axRunReq[16] THEN
		xChainInterlock := TRUE;
	END_IF

	axRunReq[12] := FALSE;		// rolki stacji 8
	axRunReq[16] := FALSE;		// rolki stacji 10

END_IF


// -------------------------------------------------------------
// BLOKADA STACJI 5 KONTRA TRANSPORTER
// -------------------------------------------------------------
//
// Wysunieta blokada znaczy "paleta ma tu stanac". Wypychanie jej
// wtedy na stacje 6 to praca transportera w zapore - i to jest
// przyczyna, dla ktorej naped 5 wchodzil w przeciazenie.
//
// WJAZD ZE STACJI 4 JEST WYJATKIEM: tam blokada MA byc wysunieta,
// bo to ona zatrzymuje palete. Dlatego warunek dotyczy wylacznie
// jazdy W STRONE STACJI 6, czyli kroku 180 toru B1.
//
// Blokada nie ma czujnika polozenia, wiec zadamy nie tylko
// zdjetej komendy, ale i tCylTime na jej faktyczne opuszczenie.
// Warunek nadrzedny, jak blokada lancucha wyzej - nie zalezy od
// tabeli krokow i zadziala takze po jej zmianie.

xSt05_BlockLock := FALSE;

IF (nOutStep = 180) AND NOT tonSt05BlockDown.Q THEN
	xSt05_BlockLock := TRUE;
	axRunReq[5] := FALSE;
	axRunReq[6] := FALSE;
END_IF


// -------------------------------------------------------------
// SPRZEZENIE: ROLKI DOCISKOWE STACJI 4 Z TRANSPORTEREM
// -------------------------------------------------------------
//
// Naped 3 (gorne rolki dociskowe) kreci sie zawsze wtedy, gdy
// kreci sie transporter stacji 4 (naped 4). Nie ma sensu, zeby
// rolki lezaly na deskach i staly, kiedy paleta pod nimi jedzie.
//
// Warunek nadrzedny, tak jak blokada lancucha wyzej: nie zalezy
// od tabeli krokow i zadziala takze po jej zmianie.
//
// Kierunek bierzemy z bitu, ktory mozna przestawic online.

axReverse[3] := xSt04_RollRev;

IF axRunReq[4] THEN
	axRunReq[3] := TRUE;
END_IF


FOR i := 1 TO cNumDrives DO

	// Naped niedopuszczony nie ruszy, chocby krok tego zadal
	IF NOT axDriveEnabled[i] THEN
		axRunReq[i] := FALSE;
	END_IF

	IF axDrvError[i] THEN
		xAnyDriveError := TRUE;
	END_IF



	// Czestotliwosc: wlasna dla napedu, inaczej bazowa.
	lrThisFreq := lrTestFreq;

	IF alrDriveFreq[i] > 0.0 THEN
		lrThisFreq := alrDriveFreq[i];
	END_IF

	// Krzywki maja wlasna nastawe i wygrywaja z tablica
	IF (i = 1) OR (i = 2) THEN
		lrThisFreq := lrCamFreq;
	END_IF

	// Naped zablokowany (blad, brak zezwolenia, zerwana
	// komunikacja) SAM kasuje u siebie zadanie ruchu - i slusznie,
	// bo nie wolno mu ruszyc samoczynnie po ustapieniu przyczyny.
	//
	// Warstwa maszyny musi wiec wydac komende OD NOWA. Dlatego:
	//   - w czasie blokady nie wolamy M_Start (byloby bez sensu,
	//     a lamaloby regule wolania na zboczu),
	//   - pamiec zbocza trzymamy wtedy wyzerowana, zeby po
	//     ustapieniu przyczyny powstalo JEDNO nowe zbocze.
	//
	// Bez tego naped, ktory raz wpadl w blad, stalby juz na
	// zawsze - skasowanie bledu nic by nie dalo, bo zbocze
	// startu dawno minelo.

	IF axRunReq[i] AND NOT axRunOld[i] AND NOT axDrvError[i] THEN
		fbNord[i].M_Start(lrFreq := lrThisFreq, xReverse := axReverse[i]);
	END_IF

	IF NOT axRunReq[i] AND axRunOld[i] THEN
		fbNord[i].M_Stop();
	END_IF

	axRunOld[i] := axRunReq[i] AND NOT axDrvError[i];

END_FOR
END_ACTION

ACTION ACT_CamCycles:
// =============================================================
// ACT_CamCycles
// Desztaplarka (st.3) i sztaplarka (st.11)
// =============================================================
//
// KORBA JEDZIE ZAWSZE W JEDNA STRONE. Cykl to jeden obrot:
// dol -> posrednia -> gorna -> DALEJ TYM SAMYM KIERUNKIEM
// z powrotem na dol. Nigdy nie wracamy tam, skad przyjechalismy.
//
// Enkoder jest jednoobrotowy i potrafi pokazac wartosc wieksza
// niz jeden obrot, wiec FB_CamAxis sprowadza ja modulo 65536,
// liczy przyrost ze znakiem i sam wykrywa przejscia przez zero.
// Tutaj operujemy juz tylko pozycjami 0..65535.
//
// REGULA NADRZEDNA obu maszyn: nic w szczekach = szczeki
// OTWARTE i jazda na pozycje DOLNA, niezaleznie od tego, gdzie
// wozek stoi.
//
// -------------------------------------------------------------
// SZCZEKI
// -------------------------------------------------------------
// KAZDY krok deklaruje xDeJawsClosed / xStJawsClosed, a cewki
// przepisujemy raz, na koncu akcji. Nie wolno polegac na tym,
// ze cewka zachowa wartosc miedzy krokami - ACT_ClearCoils
// zeruje wszystkie cewki w kazdym cyklu przy zdjetym START_TEST,
// wiec krok, ktory ich nie odswieza, traci sterowanie zaworem.
//
// -------------------------------------------------------------
// SYGNALY
// -------------------------------------------------------------
//   xPal_St03     IN2   sztapla na stacji 3
//   xPal_St04In   IN3   stacja 4 przyjela palete
//   xPal_St11     IN8   paleta na stacji 11
//
// Czujnik musi byc najpierw WOLNY, zeby sie zaliczyl.


// =============================================================
// RESET CYKLU DO ZERA
// =============================================================
//
// Wykonujemy to PRZED maszynami stanow, zeby jeszcze w tym
// samym cyklu ruszyly juz od kroku 0 - takze transport,
// bo ACT_TestFeed idzie po tej akcji.

rtrgResetCycle(CLK := RESET_CYCLE);

IF rtrgResetCycle.Q THEN

	nDeStep   := 0;
	nStStep   := 0;
	nFeedStep := 0;
	nOutStep  := 0;
	nOut2Step := 0;
	nOut3Step := 0;

	xOutStart  := FALSE;
	xOut2Start := FALSE;
	xOut3Start := FALSE;
	xSt08_RollDown  := FALSE;
	xSt08_AtStation := FALSE;

	xSt05_Done := FALSE;

	GVL_PERSIST.St03.Mem.nRemaining := 0;
	GVL_PERSIST.St03.Mem.nHeld      := 0;
	GVL_PERSIST.St11.Mem.nHeld      := 0;

	xDe_PalletReleased := FALSE;
	xSt_StackReady     := FALSE;
	xSt01_StackReady   := FALSE;

	nFeedPallets := 0;
	nDeCycles    := 0;
	nStCycles    := 0;

	RESET_CYCLE := FALSE;

END_IF


// =============================================================
// KONTROLA NASTAW POZYCJI
// =============================================================
//
// Trzy punkty musza byc od siebie oddalone o co najmniej
// diCamMinSpan, liczac najkrotsza droga po okregu. Zerowe
// nastawy - na przyklad po skasowaniu danych nieulotnych -
// znacza, ze kazdy krok od razu melduje "na pozycji", a szczeki
// zamykaja sie tam, gdzie wozek akurat stoi.

xDeCfgOK := TRUE;

diTmp := GVL_PERSIST.St03.Cfg.diPosMiddle - GVL_PERSIST.St03.Cfg.diPosBottom;
IF diTmp >  32768 THEN diTmp := diTmp - 65536; END_IF
IF diTmp < -32768 THEN diTmp := diTmp + 65536; END_IF
IF ABS(diTmp) < diCamMinSpan THEN xDeCfgOK := FALSE; END_IF

diTmp := GVL_PERSIST.St03.Cfg.diPosTop - GVL_PERSIST.St03.Cfg.diPosBottom;
IF diTmp >  32768 THEN diTmp := diTmp - 65536; END_IF
IF diTmp < -32768 THEN diTmp := diTmp + 65536; END_IF
IF ABS(diTmp) < diCamMinSpan THEN xDeCfgOK := FALSE; END_IF

diTmp := GVL_PERSIST.St03.Cfg.diPosTop - GVL_PERSIST.St03.Cfg.diPosMiddle;
IF diTmp >  32768 THEN diTmp := diTmp - 65536; END_IF
IF diTmp < -32768 THEN diTmp := diTmp + 65536; END_IF
IF ABS(diTmp) < diCamMinSpan THEN xDeCfgOK := FALSE; END_IF


xStCfgOK := TRUE;

diTmp := GVL_PERSIST.St11.Cfg.diPosMiddle - GVL_PERSIST.St11.Cfg.diPosBottom;
IF diTmp >  32768 THEN diTmp := diTmp - 65536; END_IF
IF diTmp < -32768 THEN diTmp := diTmp + 65536; END_IF
IF ABS(diTmp) < diCamMinSpan THEN xStCfgOK := FALSE; END_IF

diTmp := GVL_PERSIST.St11.Cfg.diPosTop - GVL_PERSIST.St11.Cfg.diPosBottom;
IF diTmp >  32768 THEN diTmp := diTmp - 65536; END_IF
IF diTmp < -32768 THEN diTmp := diTmp + 65536; END_IF
IF ABS(diTmp) < diCamMinSpan THEN xStCfgOK := FALSE; END_IF

diTmp := GVL_PERSIST.St11.Cfg.diPosTop - GVL_PERSIST.St11.Cfg.diPosMiddle;
IF diTmp >  32768 THEN diTmp := diTmp - 65536; END_IF
IF diTmp < -32768 THEN diTmp := diTmp + 65536; END_IF
IF ABS(diTmp) < diCamMinSpan THEN xStCfgOK := FALSE; END_IF


// =============================================================
// ZMIANA KROKU
// =============================================================
//
// Blok osi liczy xInPos wzgledem celu z POPRZEDNIEGO cyklu,
// wiec w pierwszym cyklu nowego kroku tej informacji nie
// zaliczamy - inaczej krok przeskoczylby dwa naraz.

// =============================================================
// KONTROLA ENKODERA PO STARCIE
// =============================================================
//
// Raz, w pierwszym cyklu po starcie PLC. Porownujemy odczyt
// z wartoscia zapamietana przed wylaczeniem. Roznica wieksza
// niz diEncCheckTol znaczy, ze enkoder NIE utrzymal pozycji
// i trzeba go zbazowac na dole.

IF NOT xEncCheckDone THEN

	xEncCheckDone := TRUE;

	diTmp := fbCamDestack.diPos - GVL_PERSIST.St03.Mem.diLastPos;
	IF diTmp >  32768 THEN diTmp := diTmp - 65536; END_IF
	IF diTmp < -32768 THEN diTmp := diTmp + 65536; END_IF
	diDeEncJump := diTmp;

	diTmp := fbCamStack.diPos - GVL_PERSIST.St11.Mem.diLastPos;
	IF diTmp >  32768 THEN diTmp := diTmp - 65536; END_IF
	IF diTmp < -32768 THEN diTmp := diTmp + 65536; END_IF
	diStEncJump := diTmp;

	GVL_PERSIST.St03.Mem.xNeedHoming := ABS(diDeEncJump) > diEncCheckTol;
	GVL_PERSIST.St11.Mem.xNeedHoming := ABS(diStEncJump) > diEncCheckTol;

	sEncCheck := 'enkodery utrzymaly pozycje - bazowanie zbedne';

	IF GVL_PERSIST.St03.Mem.xNeedHoming THEN
		sEncCheck := 'DESZTAPLARKA - enkoder nie utrzymal pozycji, zbazuj dol';
	END_IF

	IF GVL_PERSIST.St11.Mem.xNeedHoming THEN
		sEncCheck := 'SZTAPLARKA - enkoder nie utrzymal pozycji, zbazuj dol';
	END_IF

END_IF


// Zapamietanie biezacej pozycji na wypadek zaniku zasilania.
// PLC ma 1 s UPSa, wiec TwinCAT zdazy zapisac dane nieulotne.
GVL_PERSIST.St03.Mem.diLastPos := fbCamDestack.diPos;
GVL_PERSIST.St11.Mem.diLastPos := fbCamStack.diPos;


// Impulsy ustawienia punktu odniesienia - kasowane co cykl
xDeSetAccum := FALSE;
xStSetAccum := FALSE;


xDeNewStep := (nDeStep <> nDeStepOld);
xStNewStep := (nStStep <> nStStepOld);

nDeStepOld := nDeStep;
nStStepOld := nStStep;

IF xDeNewStep THEN
	tonDeStep(IN := FALSE);
	xDeArmed := FALSE;
END_IF

IF xStNewStep THEN
	tonStStep(IN := FALSE);
	xStArmed := FALSE;
END_IF

tonDeStep(IN := TRUE, PT := tDeStep);
tonStStep(IN := TRUE, PT := tStStep);

xDeAdvance := tonDeStep.Q AND NOT xDeNewStep;
xStAdvance := tonStStep.Q AND NOT xStNewStep;

xDeAtPos := fbCamDestack.xInPos AND NOT xDeNewStep;
xStAtPos := fbCamStack.xInPos   AND NOT xStNewStep;


// Czasowki liczone od ZACISNIECIA hamulca, nie od wejscia w krok
tonDeBrake(IN := NOT fbCamDestack.xBrakeRelease, PT := tDeBrakeWait);
tonStBrake(IN := NOT fbCamStack.xBrakeRelease,   PT := tStBrakeWait);


// =============================================================
// DESZTAPLARKA - STACJA 3
// =============================================================
//
//   0   dom: szczeki otwarte, jazda na dol
//   10  czekam na sztaple
//   20  jazda na pozycje posrednia, szczeki OTWARTE
//   30  hamulec zalozony, odliczam 1 s
//   40  szczeki zamykaja sie pod druga paleta od dolu
//   50  jazda na gore - stos uniesiony przez druga palete
//   60  info do transportu, czekam az stacja 4 przyjmie palete
//   70  DALEJ tym samym kierunkiem, dopelnienie obrotu na dol
//   80  hamulec zalozony, szczeki otwieraja sie
//   85  BRAMKA CYKLU - na dole czekam na koniec cyklu stacji 5
//   90  ostatnia paleta - nie ma czego chwytac, wyjezdza sama

xDeJog := (JOG_DESTACK_FWD OR JOG_DESTACK_REV) AND NOT START_DESTACK;

rtrgDeStart(CLK := START_DESTACK);

IF rtrgDeStart.Q THEN
	nDeStep := 0;
END_IF

IF rtrgDeStart.Q AND xAutoResetOnStart AND xAnyDriveFault THEN
	xResetInProgress := TRUE;
	nResetTries      := 0;
	xResetFailed     := FALSE;
END_IF

xDeGo        := FALSE;
tDeStep      := tJawTime;
tDeBrakeWait := tDeGripDelay;


// REGULA NADRZEDNA: pusto w szczekach w kroku niosacym stos
// to sprzecznosc - wracamy do domu zamiast jechac dalej.
IF (GVL_PERSIST.St03.Mem.nHeld <= 0) AND (nDeStep >= 50) AND (nDeStep <= 70) THEN
	nDeStep := 0;
END_IF


IF NOT START_DESTACK THEN
	sDePhase := 'DESZTAPLARKA - stop, START_DESTACK = FALSE';
END_IF

IF xDeJog THEN
	sDePhase := 'DESZT. RECZNIE - jazda krzywka, patrz na diPos';
END_IF

IF START_DESTACK AND fbCamDestack.xBrakeWait THEN
	sDePhase := 'DESZT. czekam na odpuszczenie hamulca przed startem';
END_IF

IF START_DESTACK AND fbCamDestack.xStall THEN
	sDePhase := 'DESZT. CZUWAK - falownik pracuje, a enkoder nie liczy';
END_IF

IF START_DESTACK AND fbCamDestack.xNoDrvAck THEN
	sDePhase := 'DESZT. CZUWAK - falownik 1 nie potwierdza pracy';
END_IF

IF START_DESTACK AND fbCamDestack.xStall AND axDrvFault[1] THEN
	sDePhase := 'DESZT. CZUWAK - falownik 1 w bledzie, kasuj xCmdResetDrives';
END_IF

IF START_DESTACK AND fbCamDestack.xStall AND NOT axDriveEnabled[1] THEN
	sDePhase := 'DESZT. CZUWAK - naped 1 NIEDOPUSZCZONY, ACT_Config sie nie wykonalo';
END_IF


IF START_DESTACK AND NOT xDeCfgOK THEN
	sDePhase := 'DESZT. NASTAWY POZYCJI PUSTE albo BLEDNE - naucz dol/srodek/gore';
END_IF


IF START_DESTACK AND NOT fbCamDestack.xStall AND xDeCfgOK THEN

	CASE nDeStep OF

	0:
		// REGULA NADRZEDNA: nic w szczekach = otwarte i na dol.
		//
		// Szczeki otwieramy OD RAZU, takze na gorze. Swiadomy
		// wybor: przy 1000 Nm na krzywce gorsza awaria jest
		// przeciagniecie zamknietych szczek przez stos niz
		// spadniecie palet. NIE dodawac tu zjazdu "trzymajac"
		// bez rozmowy - bylo zrobione i zostalo cofniete.
		sDePhase := 'DESZT. 0 dom: szczeki otwarte, jazda na dol';
		xDeJawsClosed := FALSE;
		GVL_PERSIST.St03.Mem.nHeld    := 0;
		xDeGo       := TRUE;
		diDeGoToEnc := GVL_PERSIST.St03.Cfg.diPosBottom;
		IF xDeAtPos THEN nDeStep := 10; END_IF

	10:
		sDePhase := 'DESZT. 1 czekam na sztaple na stacji 3 (IN2)';
		xDeJawsClosed := FALSE;
		xDe_Empty := TRUE;

		// Sztapla, ktora JUZ stoi na stacji przy wejsciu w krok,
		// jest sztapla gotowa do pracy - nie kazemy jej zjezdzac
		// i wracac. Uzbrojenie chroni tylko przed policzeniem
		// tej samej sztapli dwa razy w trakcie czekania.
		IF xDeNewStep AND xPal_St03 THEN xDeArmed := TRUE; END_IF

		IF NOT xPal_St03 THEN xDeArmed := TRUE; END_IF

		IF xDeArmed AND xPal_St03 THEN
			GVL_PERSIST.St03.Mem.nRemaining := GVL_PERSIST.St03.Cfg.nStackSize;
			xDe_Empty    := FALSE;
			nDeStep      := 20;
		END_IF

	20:
		sDePhase := 'DESZT. 2 jazda na pozycje posrednia, szczeki otwarte';
		xDeJawsClosed := FALSE;
		xDeGo       := TRUE;
		diDeGoToEnc := GVL_PERSIST.St03.Cfg.diPosMiddle;
		IF xDeAtPos THEN nDeStep := 30; END_IF

	30:
		sDePhase := 'DESZT. 3 hamulec zalozony - odliczam przed chwytem';
		xDeJawsClosed := FALSE;
		IF tonDeBrake.Q THEN nDeStep := 40; END_IF

	40:
		sDePhase := 'DESZT. 4 szczeki chwytaja 2. palete od dolu';
		xDeJawsClosed := TRUE;
		IF xDeAdvance THEN
			GVL_PERSIST.St03.Mem.nHeld := GVL_PERSIST.St03.Mem.nRemaining - 1;
			nDeStep := 50;
		END_IF

	50:
		sDePhase := 'DESZT. 5 jazda na gore - stos uniesiony';
		xDeJawsClosed := TRUE;
		xDeGo       := TRUE;
		diDeGoToEnc := GVL_PERSIST.St03.Cfg.diPosTop;
		IF xDeAtPos THEN nDeStep := 60; END_IF

	60:
		// Potwierdzeniem odbioru jest czujnik na KONCU stacji 4
		// (IN4), a nie ten od wjazdu pod rolki. Dopiero on mowi,
		// ze paleta naprawde zjechala z desztaplarki.
		//
		// TEN WARUNEK MUSI BYC KROTKI. Stos wisi tu na szczekach,
		// wiec nie wolno w tym kroku czekac na nic dalszego niz
		// zjazd palety z desztaplarki - bramka cyklu stoi w
		// kroku 85, na dole, przy stosie opartym o transporter.
		//
		// IN4 pilnuje takze tego, zeby stos nie zjechal na palete,
		// ktora jeszcze nie zdazyla wyjechac.
		sDePhase := 'DESZT. 6 paleta zwolniona - czekam na koniec st.4 (IN4)';
		xDeJawsClosed := TRUE;
		xDe_PalletReleased := TRUE;

		IF NOT xPal_St04End THEN xDeArmed := TRUE; END_IF

		IF xPal_St04End AND NOT xDeArmed THEN
			sDePhase := 'DESZT. 6 IN4 JUZ zaslonony - odslon i zaslon ponownie';
		END_IF

		IF xDeArmed AND xPal_St04End THEN
			GVL_PERSIST.St03.Mem.nRemaining       := GVL_PERSIST.St03.Mem.nRemaining - 1;
			xDe_PalletReleased := FALSE;
			nDeStep            := 70;
		END_IF

	70:
		// DALEJ tym samym kierunkiem - dopelnienie pelnego obrotu
		sDePhase := 'DESZT. 7 dopelnienie obrotu - zjazd stosu na dol';
		xDeJawsClosed := TRUE;
		xDeGo       := TRUE;
		diDeGoToEnc := GVL_PERSIST.St03.Cfg.diPosBottom;
		IF xDeAtPos THEN nDeStep := 80; END_IF

	80:
		sDePhase := 'DESZT. 8 hamulec zalozony - szczeki otwieraja sie';
		tDeBrakeWait := tJawTime;
		GVL_PERSIST.St03.Mem.nHeld := 0;

		xDeJawsClosed := TRUE;

		IF NOT fbCamDestack.xBrakeRelease THEN
			xDeJawsClosed := FALSE;
		END_IF

		IF tonDeBrake.Q AND (GVL_PERSIST.St03.Mem.nRemaining > 1) THEN
			nDeCycles := nDeCycles + 1;
			nDeStep   := 85;
		END_IF

		IF tonDeBrake.Q AND (GVL_PERSIST.St03.Mem.nRemaining = 1) THEN
			nDeCycles := nDeCycles + 1;
			nDeStep   := 90;
		END_IF

		IF tonDeBrake.Q AND (GVL_PERSIST.St03.Mem.nRemaining <= 0) THEN
			nDeStep := 0;
		END_IF

	85:
		// BRAMKA CYKLU - JEDYNE DLUGIE CZEKANIE DESZTAPLARKI.
		//
		// Stoi TU, a nie na gorze w kroku 60, i to jest istota
		// sprawy: wozek jest na dole, stos oparty o transporter,
		// szczeki otwarte, hamulec zalozony. Nic nie wisi.
		//
		// Wczesniej ta bramka stala w kroku 60 i stos zostawal
		// zawieszony na szczekach przez caly cykl stacji 5 -
		// dziesiatki sekund zamiast kilku. Tak stracilismy stos.
		//
		// Czekamy na koniec cyklu stacji 5: dopiero wtedy ma sens
		// wydawac kolejna palete, bo poprzednia zjechala juz
		// w strone stacji 16.
		sDePhase := 'DESZT. 8b stos na dole - czekam na koniec cyklu st.5';
		xDeJawsClosed := FALSE;

		IF xSt05_Done THEN
			xSt05_Done := FALSE;
			nDeStep    := 20;
		END_IF

	90:
		// Ostatnia paleta lezy wprost na transporterze - szczeki
		// nie maja pod co wejsc, wiec wyjezdza sama.
		sDePhase := 'DESZT. 9 ostatnia paleta - wyjezdza sama, bez chwytu';
		xDeJawsClosed := FALSE;
		xDe_PalletReleased := TRUE;

		IF NOT xPal_St04End THEN xDeArmed := TRUE; END_IF

		IF xPal_St04End AND NOT xDeArmed THEN
			sDePhase := 'DESZT. 9 IN4 JUZ zaslonony - odslon i zaslon ponownie';
		END_IF

		IF xDeArmed AND xPal_St04End THEN
			GVL_PERSIST.St03.Mem.nRemaining       := 0;
			xDe_PalletReleased := FALSE;
			nDeCycles          := nDeCycles + 1;
			nDeStep            := 0;
		END_IF

	END_CASE

END_IF


// =============================================================
// SZTAPLARKA - STACJA 11
// =============================================================
//
//   0   dom: szczeki otwarte, jazda na dol
//   10  czekam na pierwsza palete
//   20  hamulec zalozony, odliczam 1 s
//   25  szczeki chwytaja palete
//   30  jazda na gore - miejsce na nastepna palete
//   40  czekam na nowa palete
//   50  zjazd na srodek - stos siada na nowej palecie
//   60  hamulec zalozony, szczeki otwieraja sie
//   70  stos pelny - czekam, az zjedzie
//   80  jazda na dol pod caly stos
//   90  hamulec zalozony, odliczam 1 s
//   95  szczeki chwytaja stos od spodu

xStJog := (JOG_STACK_FWD OR JOG_STACK_REV) AND NOT START_STACK;

rtrgStStart(CLK := START_STACK);

IF rtrgStStart.Q THEN
	nStStep := 0;
END_IF

xStGo        := FALSE;
tStStep      := tJawTime;
tStBrakeWait := tDeGripDelay;


IF NOT START_STACK THEN
	sStPhase := 'SZTAPLARKA - stop, START_STACK = FALSE';
END_IF

IF xStJog THEN
	sStPhase := 'SZTAPL. RECZNIE - jazda krzywka, patrz na diPos';
END_IF

IF START_STACK AND fbCamStack.xBrakeWait THEN
	sStPhase := 'SZTAPL. czekam na odpuszczenie hamulca przed startem';
END_IF

IF START_STACK AND fbCamStack.xStall THEN
	sStPhase := 'SZTAPL. CZUWAK - falownik pracuje, a enkoder nie liczy';
END_IF

IF START_STACK AND fbCamStack.xNoDrvAck THEN
	sStPhase := 'SZTAPL. CZUWAK - falownik 2 nie potwierdza pracy';
END_IF

IF START_STACK AND fbCamStack.xStall AND axDrvFault[2] THEN
	sStPhase := 'SZTAPL. CZUWAK - falownik 2 w bledzie, kasuj xCmdResetDrives';
END_IF

IF START_STACK AND fbCamStack.xStall AND NOT axDriveEnabled[2] THEN
	sStPhase := 'SZTAPL. CZUWAK - naped 2 NIEDOPUSZCZONY, ACT_Config sie nie wykonalo';
END_IF


IF START_STACK AND NOT xStCfgOK THEN
	sStPhase := 'SZTAPL. NASTAWY POZYCJI PUSTE albo BLEDNE - naucz dol/srodek/gore';
END_IF


IF START_STACK AND NOT fbCamStack.xStall AND xStCfgOK THEN

	CASE nStStep OF

	0:
		// Szczeki otwarte od razu - patrz komentarz w kroku 0
		// desztaplarki. Swiadomy wybor.
		sStPhase := 'SZTAPL. 0 dom: szczeki otwarte, jazda na dol';
		xStJawsClosed := FALSE;
		GVL_PERSIST.St11.Mem.nHeld    := 0;
		xStGo       := TRUE;
		diStGoToEnc := GVL_PERSIST.St11.Cfg.diPosBottom;
		IF xStAtPos THEN nStStep := 10; END_IF

	10:
		sStPhase := 'SZTAPL. 1 czekam na pierwsza palete (IN8)';
		xStJawsClosed := FALSE;

		IF NOT xPal_St11 THEN xStArmed := TRUE; END_IF

		IF xPal_St11 AND NOT xStArmed THEN
			sStPhase := 'SZTAPL. 1 IN8 JUZ zaslonony - odslon i zaslon ponownie';
		END_IF

		IF xStArmed AND xPal_St11 THEN nStStep := 20; END_IF

	20:
		sStPhase := 'SZTAPL. 2 hamulec zalozony - odliczam przed chwytem';
		xStJawsClosed := FALSE;
		IF tonStBrake.Q THEN nStStep := 25; END_IF

	25:
		sStPhase := 'SZTAPL. 2b szczeki chwytaja palete';
		xStJawsClosed := TRUE;
		IF xStAdvance THEN
			GVL_PERSIST.St11.Mem.nHeld := 1;
			nStStep := 30;
		END_IF

	30:
		sStPhase := 'SZTAPL. 3 jazda na gore - miejsce na nowa palete';
		xStJawsClosed := TRUE;
		xStGo       := TRUE;
		diStGoToEnc := GVL_PERSIST.St11.Cfg.diPosTop;
		IF xStAtPos THEN nStStep := 40; END_IF

	40:
		sStPhase := 'SZTAPL. 4 czekam na nowa palete (IN8)';
		xStJawsClosed := TRUE;

		IF NOT xPal_St11 THEN xStArmed := TRUE; END_IF

		IF xPal_St11 AND NOT xStArmed THEN
			sStPhase := 'SZTAPL. 4 IN8 JUZ zaslonony - odslon i zaslon ponownie';
		END_IF

		IF xStArmed AND xPal_St11 THEN nStStep := 50; END_IF

	50:
		sStPhase := 'SZTAPL. 5 zjazd na srodek - stos siada na palecie';
		xStJawsClosed := TRUE;
		xStGo       := TRUE;
		diStGoToEnc := GVL_PERSIST.St11.Cfg.diPosMiddle;
		IF xStAtPos THEN nStStep := 60; END_IF

	60:
		sStPhase := 'SZTAPL. 6 hamulec zalozony - szczeki otwieraja sie';
		tStBrakeWait := tJawTime;

		xStJawsClosed := TRUE;

		IF NOT fbCamStack.xBrakeRelease THEN
			xStJawsClosed := FALSE;
		END_IF

		// Po inkrementacji GVL_PERSIST.St11.Mem.nHeld to liczba palet w stosie,
		// ktory lezy teraz na transporterze.
		IF tonStBrake.Q THEN
			GVL_PERSIST.St11.Mem.nHeld   := GVL_PERSIST.St11.Mem.nHeld + 1;
			nStCycles := nStCycles + 1;
			nStStep   := 80;
		END_IF

		IF tonStBrake.Q AND (GVL_PERSIST.St11.Mem.nHeld >= GVL_PERSIST.St11.Cfg.nStackSize) THEN
			nStStep := 70;
		END_IF

	70:
		sStPhase := 'SZTAPL. 7 stos pelny - czekam, az zjedzie ze stacji';
		xStJawsClosed := FALSE;
		xSt_StackReady := TRUE;

		IF NOT xPal_St11 THEN
			xSt_StackReady := FALSE;
			GVL_PERSIST.St11.Mem.nHeld        := 0;
			nStStep        := 0;
		END_IF

	80:
		sStPhase := 'SZTAPL. 8 jazda na dol - pod caly stos';
		xStJawsClosed := FALSE;
		xStGo       := TRUE;
		diStGoToEnc := GVL_PERSIST.St11.Cfg.diPosBottom;
		IF xStAtPos THEN nStStep := 90; END_IF

	90:
		sStPhase := 'SZTAPL. 9 hamulec zalozony - odliczam przed chwytem';
		xStJawsClosed := FALSE;
		IF tonStBrake.Q THEN nStStep := 95; END_IF

	95:
		sStPhase := 'SZTAPL. 9b szczeki chwytaja stos od spodu';
		xStJawsClosed := TRUE;
		IF xStAdvance THEN nStStep := 30; END_IF

	END_CASE

END_IF


// =============================================================
// POMIAR CYKLU I PRZESTAWIENIE PUNKTU ODNIESIENIA
// =============================================================
//
// Robimy to w kroku, w ktorym os STOI - nigdy w trakcie ruchu.
// Poprzednia wersja przestawiala punkt odniesienia w chwili
// dojazdu, czyli w srodku najdluzszego ruchu i wartoscia
// zalezna od enkodera. To bylo prosze o klopoty.
//
// diAccum w chwili wejscia w krok 8 to droga przejechana od
// poprzedniego dolu, czyli DLUGOSC CYKLU MASZYNY w impulsach.
// Jesli enkoder jest 1:1 z korba, wyjdzie okolo 65536.

IF xDeNewStep AND (nDeStep = 80) THEN

	diDeCycleCounts := fbCamDestack.diAccum;

	diTmp := fbCamDestack.diPos - GVL_PERSIST.St03.Cfg.diPosBottom;
	IF diTmp >  32768 THEN diTmp := diTmp - 65536; END_IF
	IF diTmp < -32768 THEN diTmp := diTmp + 65536; END_IF
	diDeBottomErr := diTmp;

	// Punkt odniesienia od zera. Wartosc nie ma juz znaczenia -
	// kazdy krok liczy swoj cel od biezacego diAccum.
	diDeAccumSet := 0;
	xDeSetAccum  := TRUE;

END_IF

IF xStNewStep AND (nStStep = 90) THEN

	diStCycleCounts := fbCamStack.diAccum;

	diTmp := fbCamStack.diPos - GVL_PERSIST.St11.Cfg.diPosBottom;
	IF diTmp >  32768 THEN diTmp := diTmp - 65536; END_IF
	IF diTmp < -32768 THEN diTmp := diTmp + 65536; END_IF
	diStBottomErr := diTmp;

	diStAccumSet := 0;
	xStSetAccum  := TRUE;

END_IF


// Najwiekszy zaobserwowany dojazd. Musi zostac MNIEJSZY niz
// diCamOvershoot - inaczej ruch do punktu tuz za nami pojedzie
// dookola calego obrotu.
//
// RESET_CAM kasuje pomiar, zeby dalo sie mierzyc od nowa bez
// pobierania projektu.

IF RESET_CAM THEN
	diDeCoastMax := 0;
	diStCoastMax := 0;
END_IF

IF ABS(fbCamDestack.diCoast) > diDeCoastMax THEN
	diDeCoastMax := ABS(fbCamDestack.diCoast);
END_IF

IF ABS(fbCamStack.diCoast) > diStCoastMax THEN
	diStCoastMax := ABS(fbCamStack.diCoast);
END_IF


// =============================================================
// DOKAD JEDZIE KROK - PRZELICZENIE RAZ, PRZY WEJSCIU
// =============================================================
//
// Krok powiedzial, do ktorej WARTOSCI ENKODERA ma dojechac.
// Tu zamieniamy to na cel na skali narastajacej, liczac droge
// do przodu z zywej pozycji - raz, w pierwszym cyklu kroku.
//
// Nigdzie nie zakladamy, ile impulsow ma cykl maszyny. Kazdy
// ruch celuje w rzeczywisty punkt na korbie, wiec blad nie ma
// sie z czego kumulowac.
//
// Jesli cel jest tuz ZA nami - mniej niz diCamOvershoot - droga
// wynosi zero. Bez tego wozek, ktory przejechal punkt o dojazd,
// objechalby caly obrot, zeby do niego wrocic.

IF xDeNewStep THEN
	diTmp := diDeGoToEnc - fbCamDestack.diPos;
	IF diTmp < 0 THEN diTmp := diTmp + 65536; END_IF
	IF diTmp >= (65536 - diCamOvershoot) THEN diTmp := 0; END_IF
	diDeTarget := fbCamDestack.diAccum + diTmp;
END_IF

IF xStNewStep THEN
	diTmp := diStGoToEnc - fbCamStack.diPos;
	IF diTmp < 0 THEN diTmp := diTmp + 65536; END_IF
	IF diTmp >= (65536 - diCamOvershoot) THEN diTmp := 0; END_IF
	diStTarget := fbCamStack.diAccum + diTmp;
END_IF


// =============================================================
// SZCZEKI -> CEWKI, CO CYKL
// =============================================================
//
// Tu i tylko tu. Kazdy krok powiedzial juz, czy szczeki maja
// byc zamkniete; my przepisujemy to na zawory w kazdym cyklu,
// zeby ACT_ClearCoils nie mogl zabrac sterowania w trakcie
// jazdy. To byl prawdziwy blad poprzedniej wersji.

IF START_DESTACK OR xDeJog THEN
	xSt03_JawClose := xDeJawsClosed;
	xSt03_JawOpen  := NOT xDeJawsClosed;
END_IF

IF START_STACK OR xStJog THEN
	xSt11_JawClose := xStJawsClosed;
	xSt11_JawOpen  := NOT xStJawsClosed;
END_IF


// =============================================================
// UCZENIE POZYCJI
// =============================================================
//
// Zbocze bitu przepisuje biezaca pozycje do nastawy. Uzywa sie
// tego przy zdjetym starcie, dojezdzajac jogiem.

rtrgTeach[1](CLK := TEACH_DE_BOTTOM);
rtrgTeach[2](CLK := TEACH_DE_MIDDLE);
rtrgTeach[3](CLK := TEACH_DE_TOP);
rtrgTeach[4](CLK := TEACH_ST_BOTTOM);
rtrgTeach[5](CLK := TEACH_ST_MIDDLE);
rtrgTeach[6](CLK := TEACH_ST_TOP);

IF rtrgTeach[1].Q THEN
	GVL_PERSIST.St03.Cfg.diPosBottom := fbCamDestack.diPos;
	sTeachLast := CONCAT('DESZT. dolna = ', DINT_TO_STRING(GVL_PERSIST.St03.Cfg.diPosBottom));
END_IF

IF rtrgTeach[2].Q THEN
	GVL_PERSIST.St03.Cfg.diPosMiddle := fbCamDestack.diPos;
	sTeachLast := CONCAT('DESZT. posrednia = ', DINT_TO_STRING(GVL_PERSIST.St03.Cfg.diPosMiddle));
END_IF

IF rtrgTeach[3].Q THEN
	GVL_PERSIST.St03.Cfg.diPosTop := fbCamDestack.diPos;
	sTeachLast := CONCAT('DESZT. gorna = ', DINT_TO_STRING(GVL_PERSIST.St03.Cfg.diPosTop));
END_IF

IF rtrgTeach[4].Q THEN
	GVL_PERSIST.St11.Cfg.diPosBottom := fbCamStack.diPos;
	sTeachLast := CONCAT('SZTAPL. dolna = ', DINT_TO_STRING(GVL_PERSIST.St11.Cfg.diPosBottom));
END_IF

IF rtrgTeach[5].Q THEN
	GVL_PERSIST.St11.Cfg.diPosMiddle := fbCamStack.diPos;
	sTeachLast := CONCAT('SZTAPL. posrednia = ', DINT_TO_STRING(GVL_PERSIST.St11.Cfg.diPosMiddle));
END_IF

IF rtrgTeach[6].Q THEN
	GVL_PERSIST.St11.Cfg.diPosTop := fbCamStack.diPos;
	sTeachLast := CONCAT('SZTAPL. gorna = ', DINT_TO_STRING(GVL_PERSIST.St11.Cfg.diPosTop));
END_IF


// =============================================================
// OSIE - JEDNO WYWOLANIE NA CYKL
// =============================================================
//
// Wolane ZAWSZE, takze przy zdjetym starcie: inaczej hamulec
// nie doliczylby swojego opoznienia po stopie, a pozycja
// przestalaby sie odswiezac na podgladzie.

fbCamDestack(
	diRawPos		:= GVL.IO_Destaker_Act_Pos,
	xEnable			:= (START_DESTACK OR xDeJog) AND xSafetyOK,
	xGoTo			:= xDeGo,
	xJogFwd			:= JOG_DESTACK_FWD AND xDeJog,
	xJogRev			:= JOG_DESTACK_REV AND xDeJog,
	diTargetAbs		:= diDeTarget,
	xSetAccum		:= xDeSetAccum,
	diSetAccumTo	:= diDeAccumSet,
	xReset			:= RESET_CAM OR rtrgResetCycle.Q,
	xDrvRunning		:= axDrvRunning[1],
	diStopLead		:= diCamStopLead,
	tBrakeReleaseLead := tCamBrakeRelease,
	tBrakeHold		:= tCamBrakeHold);

fbCamStack(
	diRawPos		:= GVL.IO_Staker_Act_Pos,
	xEnable			:= (START_STACK OR xStJog) AND xSafetyOK,
	xGoTo			:= xStGo,
	xJogFwd			:= JOG_STACK_FWD AND xStJog,
	xJogRev			:= JOG_STACK_REV AND xStJog,
	diTargetAbs		:= diStTarget,
	xSetAccum		:= xStSetAccum,
	diSetAccumTo	:= diStAccumSet,
	xReset			:= RESET_CAM OR rtrgResetCycle.Q,
	xDrvRunning		:= axDrvRunning[2],
	diStopLead		:= diCamStopLead,
	tBrakeReleaseLead := tCamBrakeRelease,
	tBrakeHold		:= tCamBrakeHold);


// -------------------------------------------------------------
// ZYCIE ENKODEROW
// -------------------------------------------------------------

IF fbCamDestack.diPos <> diDePosOld THEN
	nDeEncMoves := nDeEncMoves + 1;
	diDePosOld  := fbCamDestack.diPos;
END_IF

IF fbCamStack.diPos <> diStPosOld THEN
	nStEncMoves := nStEncMoves + 1;
	diStPosOld  := fbCamStack.diPos;
END_IF


// -------------------------------------------------------------
// ZADANIE DO WARSTWY NAPEDOW I HAMULCE
// -------------------------------------------------------------

axRunReq[1]  := fbCamDestack.xRunReq;
axReverse[1] := fbCamDestack.xRev;

axRunReq[2]  := fbCamStack.xRunReq;
axReverse[2] := fbCamStack.xRev;

xBrakeDestack := fbCamDestack.xBrakeRelease;
xBrakeStack   := fbCamStack.xBrakeRelease;
END_ACTION

ACTION ACT_ClearCoils:
// =============================================================
// ACT_ClearCoils
// Zdjecie wszystkich cewek
// =============================================================
//
// Przy zaworach dwucewkowych silownik zostaje tam, gdzie jest -
// nie wraca sam. Przy trojpolozeniowych to polozenie spoczynkowe.

xSt03_JawClose	:= FALSE;
xSt03_JawOpen	:= FALSE;

xSt04_UpExt		:= FALSE;
xSt04_UpRet		:= FALSE;
xSt04_LoExt		:= FALSE;
xSt04_LoRet		:= FALSE;

xSt05_BlockExt	:= FALSE;
xSt05_BlockRet	:= FALSE;
xSt05_LiftUp	:= FALSE;
xSt05_LiftDown	:= FALSE;
xSt05_JawClose	:= FALSE;

FOR i := 1 TO 6 DO
	axSt05_PullUp[i]	:= FALSE;
	axSt05_PullDown[i]	:= FALSE;
END_FOR

xSt08_Up		:= FALSE;
xSt08_Down		:= FALSE;
xSt10_Up		:= FALSE;
xSt10_Down		:= FALSE;

xSt11_JawClose	:= FALSE;
xSt11_JawOpen	:= FALSE;
END_ACTION

ACTION ACT_Config:
// =============================================================
// ACT_Config
// Jednorazowe ustawienia
// =============================================================

// Cala akcja wykonuje sie raz. Swiadomie BEZ instrukcji RETURN -
// w akcji programu potrafi ona wyjsc z calego POU, a wtedy nic
// dalszego by sie nie wykonalo.
IF NOT xInit THEN

xInit := TRUE;


// -------------------------------------------------------------
// DOPUSZCZENIE NAPEDOW
// -------------------------------------------------------------
//
// Domyslnie wszystkie transportery dopuszczone.

FOR i := 1 TO 20 DO
	axDriveEnabled[i] := TRUE;
END_FOR

// Krzywki podnoszenia palet. Sterowane WYLACZNIE przez
// ACT_CamCycles - tabela krokow transportu nigdy o nie nie pyta.
//   1  krzywka desztaplarki, stacja 3
//   2  krzywka sztaplarki,   stacja 11 (zasilana ze stacji 8)
axDriveEnabled[1] := TRUE;
axDriveEnabled[2] := TRUE;

// Rolki dociskowe stacji 4 - DOPUSZCZONE.
//
// Kreca sie sprzegniete z transporterem stacji 4 (naped 4):
// jedzie transporter, kreca sie rolki. Sprzezenie robi
// ACT_ApplyDrives, nie tabela krokow.
//
// Kierunek wybiera bit xSt04_RollRev, do przestawienia ONLINE.
//
// NA RAZIE ZABLOKOWANE. Przy pelnej czestotliwosci rolki pchaly
// palete tak mocno, ze wykladaly falownik transportera stacji 4.
// Rolki maja palecie TOWARZYSZYC, nie ja napedzac - ich predkosc
// obwodowa musi byc rowna predkosci transportera albo minimalnie
// nizsza.
//
// Zanim wlaczysz je z powrotem, ustaw im WLASNA czestotliwosc:
//     alrDriveFreq[3] := <Hz>
// (zero znaczy "uzyj lrTestFreq" - i to wlasnie bylo za duzo).
// Dopuszczenie: axDriveEnabled[3] := TRUE, online, bez pobierania.
axDriveEnabled[3] := FALSE;

// Falownik 20 nie istnieje w konfiguracji
axDriveEnabled[20] := FALSE;


// -------------------------------------------------------------
// KIERUNEK OBROTOW
// -------------------------------------------------------------
//
// Zle podlaczone silniki. Numery falownikow wg przydzialu:
//   stacja 1  -> falownik 8
//   stacja 3  -> falownik 10   (stwierdzone przy pierwszej probie)
//   stacja 5  -> falownik 5
//   stacja 6  -> falownik 6
//   stacja 7  -> falownik 11
//   stacja 8  -> falownik 12
//   stacja 9  -> falownik 7
//   stacja 14 -> falownik 17
//   stacja 15 -> falownik 18
//   stacja 16 -> falownik 19

FOR i := 1 TO 20 DO
	axReverse[i] := FALSE;
END_FOR

// Krzywki 1 i 2 jada w dobra strone - kierunku NIE odwracamy
// na stale. O kierunku decyduje FB_CamAxis, bo powrot do zera
// potrafi wypasc w druga strone.
axReverse[8]  := TRUE;
axReverse[10] := TRUE;		// stacja 3 - stwierdzone na maszynie
axReverse[5]  := TRUE;
axReverse[6]  := TRUE;
axReverse[11] := TRUE;
axReverse[12] := TRUE;
axReverse[7]  := TRUE;
axReverse[17] := TRUE;
axReverse[18] := TRUE;
axReverse[19] := TRUE;

END_IF
END_ACTION

ACTION ACT_Drives:
// =============================================================
// ACT_Drives
// Wywolanie falownikow - PO wystawieniu zadan
// =============================================================

xAnyDriveFault := FALSE;

FOR i := 1 TO cNumDrives DO

	fbNord[i](
		lrFmax			:= cFmax,
		xSafetyOK		:= xSafetyOK,
		// TODO: podpiac realny status EtherCAT (WcState)
		xEtherCAT_OK	:= TRUE,
		stIn			:= GVL.NORD_DRIVE_IN[i]
	);

	GVL.NORD_DRIVE_OUT[i] := fbNord[i].stOut;

	aeDrvState[i]		:= fbNord[i].eState;
	axDrvRunning[i]		:= fbNord[i].xRunning;
	axDrvFault[i]		:= fbNord[i].xFault;
	axDrvError[i]		:= fbNord[i].xError;
	awDrvStatus[i]		:= fbNord[i].wStatusWord;
	awDrvControl[i]		:= fbNord[i].wControlWord;
	alrDrvFreqAct[i]	:= fbNord[i].lrFreqActual;

	IF axDrvFault[i] THEN
		xAnyDriveFault := TRUE;
	END_IF

END_FOR
END_ACTION

ACTION ACT_Inputs:
// =============================================================
// ACT_Inputs
// Czujniki - JEDYNE miejsce, w ktorym interpretujemy polaryzacje
// =============================================================
//
// Czesc czujnikow daje 1 przy palecie, czesc 0. Nizej jest to
// sprowadzone do jednego znaczenia: xPal_* = TRUE znaczy
// PALETA JEST. Reszta programu nie zna juz polaryzacji.
//
//   IN1   stacja 1              1 = paleta   NIE UZYWANY
//   IN2   stacja 3              1 = paleta
//   IN3   za desztaplarka       0 = paleta   wjazd na stacje 4
//   IN4   koniec testu desek    0 = paleta   stacja 4
//   IN5   stacja 7              1 = paleta
//   IN6   koniec stacji 13      0 = paleta
//   IN7   stacja 8              1 = paleta
//   IN8   stacja 11             1 = paleta
//   IN9   niepodlaczony
//   IN10  stacja 16             1 = paleta


// Surowy obraz wejsc - do podgladu bez otwierania GVL
FOR i := 1 TO 10 DO
	axInRaw[i] := GVL.INPUTS[i];
END_FOR


// -------------------------------------------------------------
// POLARYZACJA - Z TABLICY, NIE Z KODU
// -------------------------------------------------------------
//
// XOR z axInInverted sprowadza kazdy czujnik do jednego
// znaczenia: TRUE = PALETA JEST. Zmiana polaryzacji to
// przestawienie jednego bitu online.

xPal_St03		:= GVL.INPUTS[2]  XOR axInInverted[2];
xPal_St04In		:= GVL.INPUTS[3]  XOR axInInverted[3];
xPal_St04End	:= GVL.INPUTS[4]  XOR axInInverted[4];
xPal_St07		:= GVL.INPUTS[5]  XOR axInInverted[5];
xPal_St13		:= GVL.INPUTS[6]  XOR axInInverted[6];
xPal_St08		:= GVL.INPUTS[7]  XOR axInInverted[7];
xPal_St11		:= GVL.INPUTS[8]  XOR axInInverted[8];
xPal_St16		:= GVL.INPUTS[10] XOR axInInverted[10];


// -------------------------------------------------------------
// STACJA 1 - BIT ZAMIAST CZUJNIKA
// -------------------------------------------------------------
//
// Czujnika IN1 swiadomie nie czytamy. Poziom xSt01_StackReady
// mowi "stos stoi i mozna nim jechac", a zbocze 0 -> 1 znaczy,
// ze na stacji 1 stanal NOWY stos.

rtrgStack(CLK := xSt01_StackReady);

IF rtrgStack.Q THEN
	nStacksSeen := nStacksSeen + 1;
END_IF
END_ACTION

ACTION ACT_Logger:
// =============================================================
// ACT_Logger
// Obserwator stanu - decyduje KIEDY pisac wiersz
// =============================================================
//
// Wiersz okresowy co tLogPeriod plus wiersz na kazde zdarzenie.
// Co JEST w wierszu - patrz ACT_LogRow. Ta akcja niczego nie
// zmienia w procesie; czyta tylko.
//
// Kolejnosc: najpierw naglowek (gdy plik dopiero powstal),
// potem ewentualny wiersz, na koncu wywolanie bloku pliku.


// -------------------------------------------------------------
// ZDARZENIA - porownanie ze stanem z poprzedniego cyklu
// -------------------------------------------------------------

xLogEvent := FALSE;
sLogWhy   := '';

// Bity, ktorych zmiana jest zdarzeniem
axLogBit[1]  := START_TEST;
axLogBit[2]  := START_FEED;
axLogBit[3]  := START_DESTACK;
axLogBit[4]  := START_STACK;
axLogBit[5]  := rtrgResetCycle.Q;
axLogBit[6]  := RESET_CAM;
axLogBit[7]  := xCmdResetDrives;
axLogBit[8]  := xSt01_StackReady;
axLogBit[9]  := xDe_PalletReleased;
axLogBit[10] := xSt05_Done;
axLogBit[11] := xSt08_PalletNOK;
axLogBit[12] := xOutStart;
axLogBit[13] := xOut2Start;
axLogBit[14] := xOut3Start;
axLogBit[15] := xDeJawsClosed;
axLogBit[16] := xStJawsClosed;
axLogBit[17] := fbCamDestack.xInPos;
axLogBit[18] := fbCamStack.xInPos;
axLogBit[19] := fbCamDestack.xStall OR fbCamDestack.xNoDrvAck;
axLogBit[20] := fbCamStack.xStall OR fbCamStack.xNoDrvAck;
axLogBit[21] := GVL_SAFETY.xSTO;
axLogBit[22] := GVL_SAFETY.xAir;
axLogBit[23] := fbCamDestack.xBrakeRelease;
axLogBit[24] := fbCamStack.xBrakeRelease;

IF NOT xLogInit THEN
	xLogInit  := TRUE;
	xLogEvent := TRUE;
	sLogWhy   := 'start';
END_IF

IF (nDeStep <> anLogStepOld[1]) OR (nStStep <> anLogStepOld[2])
   OR (nFeedStep <> anLogStepOld[3]) OR (nOutStep <> anLogStepOld[4])
   OR (nOut2Step <> anLogStepOld[5]) OR (nOut3Step <> anLogStepOld[6]) THEN
	xLogEvent := TRUE;
	sLogWhy   := CONCAT(sLogWhy, 'step ');
END_IF

FOR nLogI := 1 TO 10 DO
	IF GVL.INPUTS[nLogI] <> axLogInOld[nLogI] THEN
		xLogEvent := TRUE;
		sLogWhy   := CONCAT(sLogWhy, 'in ');
		EXIT;
	END_IF
END_FOR

FOR nLogI := 1 TO cNumDrives DO
	IF axRunReq[nLogI] <> axLogReqOld[nLogI] THEN
		xLogEvent := TRUE;
		sLogWhy   := CONCAT(sLogWhy, 'drv ');
		EXIT;
	END_IF
END_FOR

FOR nLogI := 1 TO cNumDrives DO
	IF axDrvFault[nLogI] AND NOT axLogFaultOld[nLogI] THEN
		xLogEvent := TRUE;
		sLogWhy   := CONCAT(sLogWhy, 'FAULT ');
		EXIT;
	END_IF
END_FOR

FOR nLogI := 1 TO 24 DO
	IF axLogBit[nLogI] <> axLogBitOld[nLogI] THEN
		xLogEvent := TRUE;
		sLogWhy   := CONCAT(sLogWhy, 'bit ');
		EXIT;
	END_IF
END_FOR

IF (ABS(fbCamDestack.diStep) > diLogEncJump) OR (ABS(fbCamStack.diStep) > diLogEncJump) THEN
	xLogEvent := TRUE;
	sLogWhy   := CONCAT(sLogWhy, 'ENCJUMP ');
END_IF

// Pamiec na nastepny cykl
anLogStepOld[1] := nDeStep;
anLogStepOld[2] := nStStep;
anLogStepOld[3] := nFeedStep;
anLogStepOld[4] := nOutStep;
anLogStepOld[5] := nOut2Step;
anLogStepOld[6] := nOut3Step;

FOR nLogI := 1 TO 10 DO
	axLogInOld[nLogI] := GVL.INPUTS[nLogI];
END_FOR

FOR nLogI := 1 TO cNumDrives DO
	axLogReqOld[nLogI]   := axRunReq[nLogI];
	axLogFaultOld[nLogI] := axDrvFault[nLogI];
END_FOR

FOR nLogI := 1 TO 24 DO
	axLogBitOld[nLogI] := axLogBit[nLogI];
END_FOR


// -------------------------------------------------------------
// TAKT OKRESOWY
// -------------------------------------------------------------

tonLog(IN := TRUE, PT := tLogPeriod);

IF tonLog.Q THEN
	tonLog(IN := FALSE);
	IF NOT xLogEvent THEN
		sLogWhy := 'tick';
	END_IF
	xLogEvent := TRUE;
END_IF


// -------------------------------------------------------------
// MASKI ZAWOROW FESTO - 16 cewek w jednym slowie
// -------------------------------------------------------------
//
// bit = (i-1)*2 + (j-1):  bit0 = [1,1], bit1 = [1,2], bit2 = [2,1] ...

wLogFesto1 := 0;
wLogFesto2 := 0;

FOR nLogI := 1 TO 8 DO
	FOR nLogJ := 1 TO 2 DO
		IF GVL.FestoValves_1[nLogI, nLogJ] THEN
			wLogFesto1 := wLogFesto1 OR SHL(WORD#1, (nLogI - 1) * 2 + (nLogJ - 1));
		END_IF
		IF GVL.FestoValves_2[nLogI, nLogJ] THEN
			wLogFesto2 := wLogFesto2 OR SHL(WORD#1, (nLogI - 1) * 2 + (nLogJ - 1));
		END_IF
	END_FOR
END_FOR


// -------------------------------------------------------------
// NAGLOWEK, WIERSZ, PLIK
// -------------------------------------------------------------

IF xLogEnable AND fbLog.xHeaderPending THEN
	fbLog.xHeaderMode := TRUE;
	ACT_LogRow();
	fbLog.xHeaderMode := FALSE;
END_IF

IF xLogEnable AND xLogEvent THEN
	ACT_LogRow();
	nLogRows := nLogRows + 1;
END_IF

// Nowy plik: RESET_CYCLE albo bit reczny. Bit sam sie zdejmuje.
fbLog(xNewFile := rtrgResetCycle.Q OR xLogNewFile);

xLogNewFile := FALSE;
END_ACTION

ACTION ACT_LogRow:
// =============================================================
// ACT_LogRow
// Obserwator stanu - CO jest w wierszu
// =============================================================
//
// Jedna lista kolumn dla naglowka i dla danych: metoda M_*
// dostaje nazwe i wartosc, a fbLog.xHeaderMode decyduje, ktore
// z nich trafi do pliku. Dodajesz kolumne = dopisujesz JEDNA
// linijke tutaj. Kolejnosc kolumn = kolejnosc ponizej.
//
// Nazwy kolumn krotkie i bez spacji - czyta to potem skrypt.

fbLog.M_Begin();

// -------------------------------------------------------------
// CZAS I POWOD
// -------------------------------------------------------------

fbLog.M_UInt ('t_ms',            fbLog.udiFileMs);
fbLog.M_Clock('clock');
fbLog.M_Str  ('why',             sLogWhy);
fbLog.M_UInt ('nCycles',         nCycles);


// -------------------------------------------------------------
// KROKI MASZYN STANU
// -------------------------------------------------------------

fbLog.M_Int  ('nDeStep',         nDeStep);
fbLog.M_Int  ('nStStep',         nStStep);
fbLog.M_Int  ('nFeedStep',       nFeedStep);
fbLog.M_Int  ('nOutStep',        nOutStep);
fbLog.M_Int  ('nOut2Step',       nOut2Step);
fbLog.M_Int  ('nOut3Step',       nOut3Step);
fbLog.M_Str  ('sDePhase',        sDePhase);
fbLog.M_Str  ('sFeedPhase',      sFeedPhase);
fbLog.M_Str  ('sOutPhase',       sOutPhase);


// -------------------------------------------------------------
// BITY OPERATORA I UZGODNIENIA
// -------------------------------------------------------------

fbLog.M_Bool ('START_TEST',      START_TEST);
fbLog.M_Bool ('START_FEED',      START_FEED);
fbLog.M_Bool ('START_DESTACK',   START_DESTACK);
fbLog.M_Bool ('START_STACK',     START_STACK);
fbLog.M_Bool ('RESET_CYCLE',     rtrgResetCycle.Q);
fbLog.M_Bool ('RESET_CAM',       RESET_CAM);
fbLog.M_Bool ('xCmdResetDrives', xCmdResetDrives);
fbLog.M_Bool ('xSt01_StackReady', xSt01_StackReady);
fbLog.M_Bool ('xDe_PalletReleased', xDe_PalletReleased);
fbLog.M_Bool ('xDe_Empty',       xDe_Empty);
fbLog.M_Bool ('xSt05_Done',      xSt05_Done);
fbLog.M_Bool ('xSt05_CanPass',   xSt05_CanPass);
fbLog.M_Bool ('xSt08_PalletNOK', xSt08_PalletNOK);
fbLog.M_Bool ('xSt08_AtStation', xSt08_AtStation);
fbLog.M_Bool ('xSt08_RollDown',  xSt08_RollDown);
fbLog.M_Bool ('xOutStart',       xOutStart);
fbLog.M_Bool ('xOut2Start',      xOut2Start);
fbLog.M_Bool ('xOut3Start',      xOut3Start);
fbLog.M_Bool ('xChainInterlock', xChainInterlock);
fbLog.M_Bool ('xSt05_BlockLock', xSt05_BlockLock);
fbLog.M_Bool ('xResetInProgress', xResetInProgress);
fbLog.M_Bool ('xResetFailed',    xResetFailed);
fbLog.M_Bool ('xAnyDriveFault',  xAnyDriveFault);
fbLog.M_Bool ('xAnyDriveError',  xAnyDriveError);
fbLog.M_UInt ('nFeedPallets',    nFeedPallets);
fbLog.M_UInt ('nStacksSeen',     nStacksSeen);


// -------------------------------------------------------------
// BEZPIECZENSTWO
// -------------------------------------------------------------

fbLog.M_Bool ('xSTO',            GVL_SAFETY.xSTO);
fbLog.M_Bool ('xAir',            GVL_SAFETY.xAir);
fbLog.M_Bool ('xResetCmd',       GVL_SAFETY.xResetCmd);


// -------------------------------------------------------------
// CZUJNIKI - surowe i po polaryzacji
// -------------------------------------------------------------

fbLog.M_Bool ('in1',             GVL.INPUTS[1]);
fbLog.M_Bool ('in2',             GVL.INPUTS[2]);
fbLog.M_Bool ('in3',             GVL.INPUTS[3]);
fbLog.M_Bool ('in4',             GVL.INPUTS[4]);
fbLog.M_Bool ('in5',             GVL.INPUTS[5]);
fbLog.M_Bool ('in6',             GVL.INPUTS[6]);
fbLog.M_Bool ('in7',             GVL.INPUTS[7]);
fbLog.M_Bool ('in8',             GVL.INPUTS[8]);
fbLog.M_Bool ('in9',             GVL.INPUTS[9]);
fbLog.M_Bool ('in10',            GVL.INPUTS[10]);
fbLog.M_Bool ('xPal_St03',       xPal_St03);
fbLog.M_Bool ('xPal_St04In',     xPal_St04In);
fbLog.M_Bool ('xPal_St04End',    xPal_St04End);
fbLog.M_Bool ('xPal_St07',       xPal_St07);
fbLog.M_Bool ('xPal_St13',       xPal_St13);
fbLog.M_Bool ('xPal_St08',       xPal_St08);
fbLog.M_Bool ('xPal_St11',       xPal_St11);
fbLog.M_Bool ('xPal_St16',       xPal_St16);


// -------------------------------------------------------------
// DESZTAPLARKA - stacja 3, os 1
// -------------------------------------------------------------

fbLog.M_Int  ('de_nHeld',        GVL_PERSIST.St03.Mem.nHeld);
fbLog.M_Int  ('de_nRemaining',   GVL_PERSIST.St03.Mem.nRemaining);
fbLog.M_Int  ('de_nStackSize',   GVL_PERSIST.St03.Cfg.nStackSize);
fbLog.M_UInt ('de_nCycles',      nDeCycles);
fbLog.M_Int  ('de_raw',          GVL.IO_Destaker_Act_Pos);
fbLog.M_Int  ('de_pos',          fbCamDestack.diPos);
fbLog.M_Int  ('de_accum',        fbCamDestack.diAccum);
fbLog.M_Int  ('de_remain',       fbCamDestack.diRemain);
fbLog.M_Int  ('de_step',         fbCamDestack.diStep);
fbLog.M_Int  ('de_turns',        fbCamDestack.diTurns);
fbLog.M_Int  ('de_coast',        fbCamDestack.diCoast);
fbLog.M_Int  ('de_moved',        fbCamDestack.diMoved);
fbLog.M_Int  ('de_target',       diDeTarget);
fbLog.M_Int  ('de_goToEnc',      diDeGoToEnc);
fbLog.M_Bool ('de_go',           xDeGo);
fbLog.M_Bool ('de_inPos',        fbCamDestack.xInPos);
fbLog.M_Bool ('de_atPos',        xDeAtPos);
fbLog.M_Bool ('de_runReq',       fbCamDestack.xRunReq);
fbLog.M_Bool ('de_rev',          fbCamDestack.xRev);
fbLog.M_Bool ('de_brakeRel',     fbCamDestack.xBrakeRelease);
fbLog.M_Bool ('de_brakeWait',    fbCamDestack.xBrakeWait);
fbLog.M_Bool ('de_atRest',       fbCamDestack.xAtRest);
fbLog.M_Bool ('de_stall',        fbCamDestack.xStall);
fbLog.M_Bool ('de_noDrvAck',     fbCamDestack.xNoDrvAck);
fbLog.M_Bool ('de_jawsClosed',   xDeJawsClosed);
fbLog.M_Bool ('de_armed',        xDeArmed);
fbLog.M_Bool ('de_cfgOK',        xDeCfgOK);
fbLog.M_Bool ('de_jog',          xDeJog);
fbLog.M_Int  ('de_posBottom',    GVL_PERSIST.St03.Cfg.diPosBottom);
fbLog.M_Int  ('de_posMiddle',    GVL_PERSIST.St03.Cfg.diPosMiddle);
fbLog.M_Int  ('de_posTop',       GVL_PERSIST.St03.Cfg.diPosTop);
fbLog.M_Int  ('de_cycleCounts',  diDeCycleCounts);
fbLog.M_Int  ('de_bottomErr',    diDeBottomErr);
fbLog.M_Int  ('de_coastMax',     diDeCoastMax);
fbLog.M_UInt ('de_encMoves',     nDeEncMoves);


// -------------------------------------------------------------
// SZTAPLARKA - stacja 11, os 2
// -------------------------------------------------------------

fbLog.M_Int  ('st_nHeld',        GVL_PERSIST.St11.Mem.nHeld);
fbLog.M_UInt ('st_nCycles',      nStCycles);
fbLog.M_Int  ('st_raw',          GVL.IO_Staker_Act_Pos);
fbLog.M_Int  ('st_pos',          fbCamStack.diPos);
fbLog.M_Int  ('st_accum',        fbCamStack.diAccum);
fbLog.M_Int  ('st_remain',       fbCamStack.diRemain);
fbLog.M_Int  ('st_step',         fbCamStack.diStep);
fbLog.M_Int  ('st_coast',        fbCamStack.diCoast);
fbLog.M_Int  ('st_target',       diStTarget);
fbLog.M_Int  ('st_goToEnc',      diStGoToEnc);
fbLog.M_Bool ('st_go',           xStGo);
fbLog.M_Bool ('st_inPos',        fbCamStack.xInPos);
fbLog.M_Bool ('st_runReq',       fbCamStack.xRunReq);
fbLog.M_Bool ('st_brakeRel',     fbCamStack.xBrakeRelease);
fbLog.M_Bool ('st_stall',        fbCamStack.xStall);
fbLog.M_Bool ('st_noDrvAck',     fbCamStack.xNoDrvAck);
fbLog.M_Bool ('st_jawsClosed',   xStJawsClosed);
fbLog.M_Bool ('st_armed',        xStArmed);
fbLog.M_Bool ('st_cfgOK',        xStCfgOK);
fbLog.M_Bool ('xSt_StackReady',  xSt_StackReady);


// -------------------------------------------------------------
// CEWKI - to, co poszlo na wyjscia w tym cyklu
// -------------------------------------------------------------

FOR nLogI := 1 TO 17 DO
	sLogPfx := CONCAT('out', INT_TO_STRING(nLogI));
	fbLog.M_Bool(sLogPfx, GVL.OUTPUTS[nLogI]);
END_FOR

fbLog.M_Hex  ('festo1',          wLogFesto1);
fbLog.M_Hex  ('festo2',          wLogFesto2);

fbLog.M_Bool ('xFeed05_Block',   xFeed05_Block);
fbLog.M_Bool ('xFeed05_Lift',    xFeed05_Lift);
fbLog.M_Bool ('xFeed05_Jaws',    xFeed05_Jaws);
fbLog.M_Bool ('xFeed05_Pull',    xFeed05_Pull);
fbLog.M_Bool ('xFeedPressOn',    xFeedPressOn);
fbLog.M_Bool ('xFeedPressLoOn',  xFeedPressLoOn);
fbLog.M_Bool ('xFeedRoll08Up',   xFeedRoll08Up);
fbLog.M_Bool ('xFeedRoll10Up',   xFeedRoll10Up);


// -------------------------------------------------------------
// NAPEDY 1..cNumDrives
// -------------------------------------------------------------
//
//   dN_req   zadanie z sekwencji (axRunReq)
//   dN_run   falownik potwierdza prace
//   dN_flt   blad falownika (bit 3 StatusWord)
//   dN_sw    StatusWord szesnastkowo
//   dN_st    stan bloku FB_NordSK550PP (E_NordSK550P_State)
//   dN_hz    czestotliwosc rzeczywista

FOR nLogI := 1 TO cNumDrives DO
	sLogPfx := CONCAT('d', INT_TO_STRING(nLogI));
	fbLog.M_Bool(CONCAT(sLogPfx, '_req'), axRunReq[nLogI]);
	fbLog.M_Bool(CONCAT(sLogPfx, '_run'), axDrvRunning[nLogI]);
	fbLog.M_Bool(CONCAT(sLogPfx, '_flt'), axDrvFault[nLogI]);
	fbLog.M_Hex (CONCAT(sLogPfx, '_sw'),  UINT_TO_WORD(awDrvStatus[nLogI]));
	fbLog.M_Int (CONCAT(sLogPfx, '_st'),  TO_DINT(aeDrvState[nLogI]));
	fbLog.M_Real(CONCAT(sLogPfx, '_hz'),  alrDrvFreqAct[nLogI]);
END_FOR


// -------------------------------------------------------------
// SAM LOGGER - zeby bylo widac, czy nie gubi
// -------------------------------------------------------------

fbLog.M_UInt ('log_dropped',     fbLog.nLinesDropped);
fbLog.M_UInt ('log_errors',      fbLog.nErrors);
fbLog.M_UInt ('log_lastErr',     fbLog.nLastErrId);

fbLog.M_End();
END_ACTION

ACTION ACT_ManualCyl:
// =============================================================
// ACT_ManualCyl
// Reczne sterowanie jednym silownikiem
// =============================================================
//
// Sluzy do sprawdzenia, czy dane wyjscie w ogole dochodzi do
// zaworu. Sekwencja stoi, transportery stoja - rusza sie tylko
// to, co wybierzesz.
//
// xManExtend i xManRetract dzialaja poziomem, nie zboczem:
// trzymasz bit, cewka jest podana.

ACT_ClearCoils();

IF NOT xManExtend AND NOT xManRetract THEN
	sPhase := CONCAT('RECZNIE - silownik ', INT_TO_STRING(nManCyl));
	sPhase := CONCAT(sPhase, ' - brak komendy');
	RETURN;
END_IF

IF xManExtend AND xManRetract THEN
	sPhase := 'RECZNIE - obie komendy naraz, nic nie robie';
	RETURN;
END_IF


sPhase := CONCAT('RECZNIE - silownik ', INT_TO_STRING(nManCyl));


CASE nManCyl OF

1:	xSt03_JawClose	:= xManExtend;
	xSt03_JawOpen	:= xManRetract;

2:	xSt04_UpExt		:= xManExtend;
	xSt04_UpRet		:= xManRetract;

3:	xSt04_LoExt		:= xManExtend;
	xSt04_LoRet		:= xManRetract;

4:	xSt05_BlockExt	:= xManExtend;
	xSt05_BlockRet	:= xManRetract;

5:	xSt05_LiftUp	:= xManExtend;
	xSt05_LiftDown	:= xManRetract;

6:	xSt05_JawClose	:= xManExtend;

7:	axSt05_PullUp[1]	:= xManExtend;
	axSt05_PullDown[1]	:= xManRetract;

8:	axSt05_PullUp[2]	:= xManExtend;
	axSt05_PullDown[2]	:= xManRetract;

9:	axSt05_PullUp[3]	:= xManExtend;
	axSt05_PullDown[3]	:= xManRetract;

10:	axSt05_PullUp[4]	:= xManExtend;
	axSt05_PullDown[4]	:= xManRetract;

11:	axSt05_PullUp[5]	:= xManExtend;
	axSt05_PullDown[5]	:= xManRetract;

12:	axSt05_PullUp[6]	:= xManExtend;
	axSt05_PullDown[6]	:= xManRetract;

13:	xSt08_Up		:= xManExtend;
	xSt08_Down		:= xManRetract;

14:	xSt10_Up		:= xManExtend;
	xSt10_Down		:= xManRetract;

15:	xSt11_JawClose	:= xManExtend;
	xSt11_JawOpen	:= xManRetract;

ELSE
	sPhase := 'RECZNIE - nieznany numer silownika';

END_CASE
END_ACTION

ACTION ACT_Move:
// =============================================================
// ACT_Move
// Przejazd miedzy stacjami - mechanika stoi
// =============================================================
//
// Pracuje PARA transporterow: ten, z ktorego paleta zjezdza,
// i ten, na ktory wjezdza. Wyjatkiem jest przejazd poprzeczny,
// gdzie jedzie sam lancuch.

tThisStep := tStepTime;

// TRUE = przejazd ma jeszcze kroki wewnetrzne, nIdx zostaje
xHoldIdx := FALSE;


CASE nIdx OF

1:	axRunReq[8] := TRUE;  axRunReq[9] := TRUE;
	sPhase := 'przejazd st.1 -> st.2   (falowniki 8 + 9)';

2:	axRunReq[9] := TRUE;  axRunReq[10] := TRUE;
	xWaitSensor := TRUE;  xSensorOK := xPal_St03;
	sPhase := 'przejazd st.2 -> st.3, czekam na czujnik st.3 (IN2)';

3:	ACT_MoveSt04();

4:	axRunReq[4] := TRUE;  axRunReq[5] := TRUE;
	sPhase := 'przejazd st.4 -> st.5   (falowniki 4 + 5)';

5:	axRunReq[5] := TRUE;  axRunReq[6] := TRUE;
	sPhase := 'przejazd st.5 -> st.6   (falowniki 5 + 6)';

6:	axRunReq[6] := TRUE;  axRunReq[11] := TRUE;
	xWaitSensor := TRUE;  xSensorOK := xPal_St07;
	sPhase := 'przejazd st.6 -> st.7, czekam na czujnik st.7 (IN5)';

7:	axRunReq[11] := TRUE; axRunReq[12] := TRUE;
	xWaitSensor := TRUE;  xSensorOK := xPal_St08;
	sPhase := 'przejazd st.7 -> st.8, czekam na czujnik st.8 (IN7)';

8:	axRunReq[12] := TRUE; axRunReq[13] := TRUE;
	xWaitSensor := TRUE;  xSensorOK := xPal_St11;
	sPhase := 'przejazd st.8 -> st.11, czekam na czujnik st.11 (IN8)';

9:	axRunReq[13] := TRUE; axRunReq[14] := TRUE;
	sPhase := 'przejazd st.11 -> st.12 (falowniki 13 + 14)';

10:	axRunReq[14] := TRUE; axRunReq[15] := TRUE;
	xWaitSensor := TRUE;  xSensorOK := xPal_St13;
	sPhase := 'przejazd st.12 -> st.13, czekam na czujnik st.13 (IN6)';

12:	// Przejazd poprzeczny. Rolki stacji 8 i 10 sa opuszczone,
	// paleta lezy na lancuchu - te transportery MUSZA stac.
	axRunReq[7] := TRUE;
	tThisStep := tChainTime;
	sPhase := 'przejazd st.8 -> st.10 lancuchem (falownik 7)';

13:	axRunReq[16] := TRUE; axRunReq[17] := TRUE;
	sPhase := 'przejazd st.10 -> st.14 (falowniki 16 + 17)';

14:	axRunReq[17] := TRUE; axRunReq[18] := TRUE;
	sPhase := 'przejazd st.14 -> st.15 (falowniki 17 + 18)';

15:	axRunReq[18] := TRUE; axRunReq[19] := TRUE;
	xWaitSensor := TRUE;  xSensorOK := xPal_St16;
	sPhase := 'przejazd st.15 -> st.16, czekam na czujnik st.16 (IN10)';

ELSE
	sPhase := 'przejazd poza tabela';

END_CASE


// Po przejezdzie paleta stoi na nastepnej stacji.
// xHoldIdx znaczy, ze przejazd ma jeszcze wlasne kroki wewnetrzne
// (stacja 4) - wtedy nIdx zostaje, przesuwa sie samo nSub.

IF xAdvance AND NOT xHoldIdx THEN
	nIdx	:= nIdx + 1;
	nSub	:= 0;
	xMoving	:= FALSE;

	IF nIdx > cLastIdx THEN
		nIdx := 0;
	END_IF
END_IF
END_ACTION

ACTION ACT_MoveSt04:
// =============================================================
// ACT_MoveSt04
// Przejazd st.3 -> st.4 z testem wytrzymalosci desek
// =============================================================
//
// Stacja 4 bada JADACA palete - transporter nie staje pod
// rolkami. Przebieg:
//
//   0   jedziemy, czekamy na czujnik wjazdu IN3
//   10  odstep tSt04_EntryToPress, zeby paleta weszla pod rolki
//   20  schodza dociski GORNE
//   30  dochodza DOLNE (tSt04_UpToLo pozniej), trwa test,
//       czekamy na czujnik konca testu IN4
//   40  dociski cofniete, paleta dojezdza tSt04_StopDelay i stoi
//
// Falownik 3 (same rolki dociskowe) jest zablokowany w
// axDriveEnabled - to nie jest transporter.

// Transportery obu stacji jada przez CALY test. Paleta jest
// dluga i przy wjezdzie lezy jeszcze na stacji 3.
axRunReq[10] := TRUE;
axRunReq[4]  := TRUE;

// Domyslnie krok jest wewnetrzny - nIdx zostaje na 3
xHoldIdx := TRUE;


CASE nSub OF

	0:
		sPhase := 'st.3->4 jazda, czekam na czujnik wjazdu (IN3)';
		xWaitSensor := TRUE;
		xSensorOK   := xPal_St04In;
		IF xAdvance THEN nSub := 10; END_IF

	10:
		sPhase := 'st.4 paleta wchodzi pod rolki - odstep';
		tThisStep := tSt04_EntryToPress;
		IF xAdvance THEN nSub := 20; END_IF

	20:
		sPhase := 'st.4 dociski gorne schodza na deski';
		xSt04_UpExt := TRUE;	xSt04_UpRet := FALSE;
		tThisStep := tSt04_UpToLo;
		IF xAdvance THEN nSub := 30; END_IF

	30:
		sPhase := 'st.4 TEST - czekam na czujnik konca testu (IN4)';
		xSt04_UpExt := TRUE;	xSt04_UpRet := FALSE;
		xSt04_LoExt := TRUE;	xSt04_LoRet := FALSE;
		xWaitSensor := TRUE;
		xSensorOK   := xPal_St04End;
		IF xAdvance THEN nSub := 40; END_IF

	40:
		sPhase := 'st.4 koniec testu - dociski cofniete, dojazd';
		xSt04_UpExt := FALSE;	xSt04_UpRet := TRUE;
		xSt04_LoExt := FALSE;	xSt04_LoRet := TRUE;
		tThisStep := tSt04_StopDelay;
		xHoldIdx  := FALSE;

END_CASE


// Bezpiecznik: czujnik konca testu zdejmuje dociski od razu,
// nie czekajac na przejscie kroku. Rolki nie maja prawa jechac
// dalej po palecie, ktora juz wyszla spod nich.
IF xPal_St04End AND (nSub = 30) THEN
	xSt04_UpExt := FALSE;	xSt04_UpRet := TRUE;
	xSt04_LoExt := FALSE;	xSt04_LoRet := TRUE;
END_IF
END_ACTION

ACTION ACT_Outputs:
// =============================================================
// ACT_Outputs
// Cewki -> wyjscia
// =============================================================
//
// CALE mapowanie zaworow siedzi tutaj i tylko tutaj. Jesli
// ktores przypisanie okaze sie odwrotne, poprawka jest w jednej
// linii, a nie w sekwencji.
//
// xCylEnable = FALSE zdejmuje cewki cylindrow linii - wtedy
// test sprawdza same transportery.
//
// NIE dziala jednak wtedy, gdy pracuje ktoras krzywka. Szczeki
// sztaplarki i desztaplarki trzymaja wtedy stos, a zdjecie ich
// cewek razem z reszta po prostu by go upuscilo.

IF NOT xCylEnable AND NOT START_DESTACK AND NOT START_STACK THEN
	ACT_ClearCoils();
END_IF


// -------------------------------------------------------------
// STACJA 3 - SZCZEKI DESZTAPLARKI
// -------------------------------------------------------------

GVL.OUTPUTS[14]	:= xSt03_JawClose;		// zamykanie
GVL.OUTPUTS[15]	:= xSt03_JawOpen;		// otwieranie


// -------------------------------------------------------------
// STACJA 4 - DOCISKI
// -------------------------------------------------------------
//
// Obie grupy gornych chodza razem: [7]/[2] to zewnetrzne
// i srodkowa, [5]/[6] to srodkowe.

GVL.OUTPUTS[7]	:= xSt04_UpExt;
GVL.OUTPUTS[2]	:= xSt04_UpRet;
GVL.OUTPUTS[5]	:= xSt04_UpExt;
GVL.OUTPUTS[6]	:= xSt04_UpRet;

GVL.OUTPUTS[4]	:= xSt04_LoExt;
GVL.OUTPUTS[3]	:= xSt04_LoRet;


// -------------------------------------------------------------
// STACJA 5
// -------------------------------------------------------------
//
// [7,2] wysuwanie blokady, [7,1] opuszczanie blokady
// [6,2] podnoszenie szczek, [6,1] opuszczanie szczek
// [1..3,1] TRUE = szczeki zamkniete

GVL.FestoValves_1[7,2]	:= xSt05_BlockExt;
GVL.FestoValves_1[7,1]	:= xSt05_BlockRet;

GVL.FestoValves_1[6,2]	:= xSt05_LiftUp;
GVL.FestoValves_1[6,1]	:= xSt05_LiftDown;

GVL.FestoValves_1[1,1]	:= xSt05_JawClose;
GVL.FestoValves_1[2,1]	:= xSt05_JawClose;
GVL.FestoValves_1[3,1]	:= xSt05_JawClose;


// Silowniki rozrywajace. NUMER ZAWORU NIE JEST NUMEREM
// SILOWNIKA - stad ta tabela zamiast petli.
GVL.FestoValves_2[4,2]	:= axSt05_PullUp[1];
GVL.FestoValves_2[4,1]	:= axSt05_PullDown[1];
GVL.FestoValves_2[3,2]	:= axSt05_PullUp[2];
GVL.FestoValves_2[3,1]	:= axSt05_PullDown[2];
GVL.FestoValves_2[1,2]	:= axSt05_PullUp[3];
GVL.FestoValves_2[1,1]	:= axSt05_PullDown[3];
GVL.FestoValves_2[2,2]	:= axSt05_PullUp[4];
GVL.FestoValves_2[2,1]	:= axSt05_PullDown[4];
GVL.FestoValves_2[5,2]	:= axSt05_PullUp[5];
GVL.FestoValves_2[5,1]	:= axSt05_PullDown[5];
GVL.FestoValves_2[6,2]	:= axSt05_PullUp[6];
GVL.FestoValves_2[6,1]	:= axSt05_PullDown[6];


// -------------------------------------------------------------
// ROLKI PODNOSZONE
// -------------------------------------------------------------

GVL.OUTPUTS[11]	:= xSt08_Up;
GVL.OUTPUTS[13]	:= xSt08_Down;
GVL.OUTPUTS[10]	:= xSt10_Up;
GVL.OUTPUTS[12]	:= xSt10_Down;


// -------------------------------------------------------------
// STACJA 11 - SZCZEKI SZTAPLARKI
// -------------------------------------------------------------

GVL.OUTPUTS[9]	:= xSt11_JawClose;
GVL.OUTPUTS[8]	:= xSt11_JawOpen;


// -------------------------------------------------------------
// HAMULCE KRZYWEK
// -------------------------------------------------------------
//
// TRUE = hamulec ROZLACZONY, mozna jechac.
// FALSE = hamulec ZALOZONY - i taki jest stan bez zasilania,
// wiec zanik napiecia trzyma wozek, a nie go puszcza.
//
// Opoznienie zalozenia (1 s 900 ms po bicie stopu) siedzi
// w FB_CamAxis - silnik hamuje wlasna rampa 2 s.

GVL.OUTPUTS[16]	:= xBrakeDestack;
GVL.OUTPUTS[17]	:= xBrakeStack;


// -------------------------------------------------------------
// DOWOD, ZE TO SIE WYKONALO
// -------------------------------------------------------------

nOutWrites := nOutWrites + 1;

nCoilsOn := 0;

IF GVL.OUTPUTS[2]  THEN nCoilsOn := nCoilsOn + 1; END_IF
IF GVL.OUTPUTS[3]  THEN nCoilsOn := nCoilsOn + 1; END_IF
IF GVL.OUTPUTS[4]  THEN nCoilsOn := nCoilsOn + 1; END_IF
IF GVL.OUTPUTS[5]  THEN nCoilsOn := nCoilsOn + 1; END_IF
IF GVL.OUTPUTS[6]  THEN nCoilsOn := nCoilsOn + 1; END_IF
IF GVL.OUTPUTS[7]  THEN nCoilsOn := nCoilsOn + 1; END_IF
IF GVL.OUTPUTS[8]  THEN nCoilsOn := nCoilsOn + 1; END_IF
IF GVL.OUTPUTS[9]  THEN nCoilsOn := nCoilsOn + 1; END_IF
IF GVL.OUTPUTS[10] THEN nCoilsOn := nCoilsOn + 1; END_IF
IF GVL.OUTPUTS[11] THEN nCoilsOn := nCoilsOn + 1; END_IF
IF GVL.OUTPUTS[12] THEN nCoilsOn := nCoilsOn + 1; END_IF
IF GVL.OUTPUTS[13] THEN nCoilsOn := nCoilsOn + 1; END_IF
IF GVL.OUTPUTS[14] THEN nCoilsOn := nCoilsOn + 1; END_IF
IF GVL.OUTPUTS[15] THEN nCoilsOn := nCoilsOn + 1; END_IF
IF GVL.OUTPUTS[16] THEN nCoilsOn := nCoilsOn + 1; END_IF
IF GVL.OUTPUTS[17] THEN nCoilsOn := nCoilsOn + 1; END_IF

FOR i := 1 TO 8 DO
	IF GVL.FestoValves_1[i,1] THEN nCoilsOn := nCoilsOn + 1; END_IF
	IF GVL.FestoValves_1[i,2] THEN nCoilsOn := nCoilsOn + 1; END_IF
	IF GVL.FestoValves_2[i,1] THEN nCoilsOn := nCoilsOn + 1; END_IF
	IF GVL.FestoValves_2[i,2] THEN nCoilsOn := nCoilsOn + 1; END_IF
END_FOR
END_ACTION

